// TIA Portal project "test_done_13_5" (V17)
// Vorlageprojekt für das Buch mit Zielsystem S7-1200

(* hardware
DEVICE "S71500/ET200MP station_1"  S7-1500 station
   slot 0: "Rail_0"  Rack  6ES7 590-1***0-0AA0
   slot 1: "PLC_2"  CPU 1516-3 PN/DP  6ES7 516-3AN02-0AB0  V2.8
      slot 3: "CPU display_1"  6ES7591-1BA00-0AA0
      slot 32768: "PROFINET interface_1"  X1
         slot 32769: "Port_1"  X1 P1
         slot 32770: "Port_2"  X1 P2
      slot 33024: "PROFINET interface_2"  X2
      slot 33280: "DP interface_1"  X3
      slot 34817: "Virtual CP interface port_1"  Virtual CP interface port  Virtual CP interface port
*)

// ===== PLC "PLC_2"  CPU 1516-3 PN/DP =====

VAR_GLOBAL CONSTANT   // PLC tag table "Standard-Variablentabelle"
   "Keiner" : Pip := 65535;
   "Automatische Aktualisierung" : Pip := 0;
   "TPA 1" : Pip := 1;
   "TPA 2" : Pip := 2;
   "TPA 3" : Pip := 3;
   "TPA 4" : Pip := 4;
   "TPA OB Servo" : Pip := 32768;
   "Local~MC(1)" : Hw_SubModule := 51;
   "Local~Common(1)" : Hw_SubModule := 50;
   "Local~Device(1)" : Hw_Device := 32;
   "Local~Configuration(1)" : Hw_SubModule := 33;
   "Local~Exec(1)" : Hw_SubModule := 52;
   "Local(1)" : Hw_SubModule := 49;
   "Local~PROFINET-Schnittstelle_1" : Hw_Interface := 64;
   "Local~PROFINET-Schnittstelle_1~Port_1" : Hw_Interface := 65;
   "Local~HSC_1(1)" : Hw_Hsc := 257;
   "Local~HSC_2(1)" : Hw_Hsc := 258;
   "Local~HSC_3(1)" : Hw_Hsc := 259;
   "Local~HSC_4(1)" : Hw_Hsc := 260;
   "Local~HSC_5(1)" : Hw_Hsc := 261;
   "Local~HSC_6(1)" : Hw_Hsc := 262;
   "Local~AI_2_1" : Hw_SubModule := 263;
   "Local~DI_6_DQ_4_1" : Hw_SubModule := 264;
   "Local~Pulse_1(1)" : Hw_Pwm := 265;
   "Local~Pulse_2(1)" : Hw_Pwm := 266;
   "Local~Pulse_3(1)" : Hw_Pwm := 267;
   "Local~Pulse_4(1)" : Hw_Pwm := 268;
   "OB_Main(1)" : OB_PCYCLE := 1;
END_VAR

VAR_GLOBAL   // PLC tag table "TAGS"
   "Start" AT %I0.0 : Bool;   // Nút nhấn start
   "Stop" AT %I0.1 : Bool;   // Nút nhấn stop
   "Nhap hang" AT %I0.2 : Bool;   // Nút nhấn nhập hàng
   "Xuat hang" AT %I0.3 : Bool;   // Nút nhấn xuất hàng
   "Nut tang" AT %I0.4 : Bool;   // nút nhấn tăng vị trí
   "Nut giam" AT %I0.5 : Bool;   // nút nhấn giảm vị trí
   "CB vi tri nhan hang" AT %I0.6 : Bool;   // cảm biến vị trí nhận hàng
   "CB vi tri xuat hang" AT %I0.7 : Bool;   // cảm biến vị trí xuất hàng
   "CB hang da xuat" AT %I1.0 : Bool;   // cảm biến báo hàng đã xuất
   "CB ban nang VT giua" AT %I1.1 : Bool;   // cảm biến bàn nâng ở vị trí giữa
   "CB ban nang VT phai" AT %I1.2 : Bool;   // cảm biến bàn nâng ở vị trí phải
   "CB ban nang VT Trai" AT %I1.3 : Bool;   // cảm biến bàn nâng ở vị trí trái
   "CB vi tri nhap hang" AT %I1.4 : Bool;   // cảm biến vị trí nhập hàng
   "Ban nang dang moving x" AT %I1.5 : Bool;   // bit báo bàn nâng đang di chuyển theo trục x
   "Ban nang dang moving z" AT %I1.6 : Bool;   // bit báo bàn nâng đang di chuyển theo trục z
   "Q_Den_Run" AT %Q0.0 : Bool;   // đầu ra - đèn run
   "Q_Ban_Nang_Nang_len" AT %Q0.1 : Bool;   // đầu ra - bàn nâng nâng lên
   "Q_ban nang sang phai" AT %Q0.2 : Bool;   // đầu ra - bàn nâng sang phải
   "Q ban nang sang trai" AT %Q0.3 : Bool;   // đầu ra - bàn nâng sang trái
   "Q bang tai nhap hang1" AT %Q0.4 : Bool;   // đầu ra - băng tải nhập hàng 1
   "Q bang tai nhap hang 2" AT %Q0.5 : Bool;   // đầu ra - băng tải nhập hàng 2
   "Q bang tai xuat hang 1" AT %Q0.6 : Bool;   // đầy ra - băng tải xuất hàng 1
   "Q bang tai xuat hang 2" AT %Q0.7 : Bool;   // đầu ra - băng tải xuất hàng 2
   "Cai vi tri nhap xuat hang" AT %QD34 : DInt;   // đầu ra - vị trí cần nhập xuất hàng
   "Hien thi vi tri nhap xuat hang" AT %QD38 : DInt;   // đầu ra - hiển thị vị trí đã chọn để nhập xuất hàng
END_VAR

VAR_GLOBAL   // PLC tag table "XUNG P"
   "P1" AT %M10.0 : Bool;
   "P2" AT %M10.1 : Bool;
   "P3" AT %M10.2 : Bool;
   "P4" AT %M10.3 : Bool;
   "P5" AT %M10.4 : Bool;
   "P6" AT %M10.5 : Bool;
   "P7" AT %M10.6 : Bool;
   "P8" AT %M10.7 : Bool;
   "P9" AT %M11.0 : Bool;
   "P10" AT %M11.1 : Bool;
   "P11" AT %M11.2 : Bool;
   "P12" AT %M11.3 : Bool;
   "P13" AT %M11.4 : Bool;
   "P14" AT %M11.5 : Bool;
   "P15" AT %M11.6 : Bool;
   "P16" AT %M11.7 : Bool;
   "P17" AT %M12.0 : Bool;
   "P18" AT %M12.1 : Bool;
   "P19" AT %M12.2 : Bool;
   "P20" AT %M12.3 : Bool;
END_VAR

VAR_GLOBAL   // PLC tag table "TRUNG GIAN"
   "Dang nhap hang" AT %M20.0 : Bool;
   "Dang xuat hang" AT %M20.1 : Bool;
   "Nhap hang - Buoc 1: Chay BT1,2" AT %M20.2 : Bool;
   "Nhap hang - Buoc 2: Lay hang" AT %M20.3 : Bool;
   "Nhap hang - Buoc 3: Dua hang vao vi tri" AT %M20.4 : Bool;
   "Nhap hang - Buoc 4: Ve vi tri home" AT %M20.5 : Bool;
   "TG_CB_VT_Nhan_Hang" AT %M20.6 : Bool;
   "TG_nhap_hang_buoc3" AT %M20.7 : Bool;
   "Xuat hang - Buoc 1: Di chuyen den vi tri lay" AT %M21.0 : Bool;
   "Xuat hang - Buoc 2: Lay hang" AT %M21.1 : Bool;
   "TG_xuat_hang_buoc2" AT %M21.2 : Bool;
   "Xuat hang - Buoc 3: Ve vi tri home" AT %M21.3 : Bool;
   "TG_xuat_hang_buoc3" AT %M21.4 : Bool;
   "Xuat hang - Buoc 4: BT chuyen hang di" AT %M21.5 : Bool;
   "TG_CB hang da xuat" AT %M21.6 : Bool;
   "TG_xuat_hang_buoc4" AT %M21.7 : Bool;
END_VAR

VAR_GLOBAL   // PLC tag table "TAGS MQTT"
   "MQTT_AutoEnable" AT %M30.0 : Bool;   // Luôn Enable MQTT Protocol
   "MQTT_AutoSubscribe" AT %M30.1 : Bool;
   "MQTT_Publish_Trigger" AT %M30.3 : Bool;
   "MQTT_Subscribe_Trigger" AT %M30.4 : Bool;
   "MQTT_Unsubscribe_Trigger" AT %M30.5 : Bool;
   "MQTT_Subscribe_P" AT %M30.6 : Bool;
   "Disable" AT %M30.7 : Bool;
   "Temp" AT %M31.0 : Bool;
END_VAR

// folder: Common

TYPE "typeDiagnostics"
TITLE = typeDiagnostics
// Provides a structure for detailed diagnostics
   STRUCT
      status : Word;   // Status of the block or error identification when error occurred
      subfunctionStatus : DWord;   // Status or return value of called FBs, FCs and system blocks
      stateNumber : DInt;   // State in the state machine of the block where the error occurred
   END_STRUCT;
END_TYPE

// folder: MqttClient

TYPE "MqttPublishPacket"
   STRUCT
      DUP_flag : Bool;
      QoS_level : Int;
      Retain : Bool;
      PublishTopic : String;
      PublishMessage : String;
   END_STRUCT;
END_TYPE

TYPE "MqttSubscribePacket"
   STRUCT
      TopicFilter : Array[0..9] of String;
      RequestedQoS : Array[0..9] of Byte;
   END_STRUCT;
END_TYPE

TYPE "MqttUnsubscribePacket"
   STRUCT
      TopicFilter : Array[0..9] of String;
   END_STRUCT;
END_TYPE

TYPE "MqttConnectPacket"
   STRUCT
      cleanSession : Bool := True;
      willFlag : Bool;
      willQoS_level : Int;
      willRetain : Bool;   // must be false, if Will flag is false
      passwordFlag : Bool := false;   // if true, a password is required
      userNameFlag : Bool := false;   // if true, a username is required
      keepAliveTime : Word := 10;
      clientIdentifier : String[23] := 'mqttdemo';
      willTopic : String[100] := 'myWill';
      willMessage : String[100] := 'This is my Will message';
      userName : String[20] := '';
      password : String[20] := '';
   END_STRUCT;
END_TYPE

// folder: (top level)

DATA_BLOCK "DB_WMS_Interface"   // DB17
{ S7_Optimized_Access := 'FALSE' }
VERSION : 0.1
   VAR
      Control_From_HMI : Struct
         Nhap_hang : Bool;
         Xuat_hang : Bool;
         Nut_tang : Bool;
         Nut_giam : Bool;
         Start : Bool;
         Stop : Bool;
         Cmd_Store_A01 : Bool;
         Cmd_Store_A02 : Bool;
         Cmd_Store_A03 : Bool;
         Cmd_Retrieve : Bool;
         Cmd_Reset : Bool;
      END_STRUCT;
      System_Feedback : Struct
         CB_vi_tri_nhan : Bool;
         CB_vi_tri_xuat : Bool;
         Moving_X : Bool;
         Moving_Z : Bool;
         Q_Den_Run : Bool;
      END_STRUCT;
      Warehouse_Data : Struct
         Cai_vi_tri_nhap_xuat : DInt;
         Hien_thi_vi_tri_nhap_xuat : DInt;
      END_STRUCT;
   END_VAR
BEGIN
END_DATA_BLOCK

DATA_BLOCK "MQTT_Client_DB"   // DB18
{ S7_Optimized_Access := 'TRUE' }
AUTHOR : YU_WEN_TANG
FAMILY : SLT_APC_FA
NAME : SLTAPCFA_1
VERSION : 1.0
// stored: InstanceOfName MQTT_Client
"MQTT_Client"
BEGIN
END_DATA_BLOCK

DATA_BLOCK "MqttControlPacket"   // DB19
{ S7_Optimized_Access := 'TRUE' }
VERSION : 0.1
   VAR
      ConnectPacket : "MqttConnectPacket";
      PublishPacket : "MqttPublishPacket";
      SubscribePacket : "MqttSubscribePacket";
      UnsubscribePacket : "MqttUnsubscribePacket";
   END_VAR
BEGIN
   SubscribePacket.TopicFilter[0] := 'factoryio/warehouse/cmd/system';
   PublishPacket.PublishTopic := 'factoryio/warehouse/bin_status';
   SubscribePacket.TopicFilter[1] := 'factoryio/warehouse/cmd/store';
   SubscribePacket.TopicFilter[2] := 'factoryio/warehouse/cmd/retrieve';
END_DATA_BLOCK

DATA_BLOCK "FB_Parse_MQTT_DB"   // DB20
{ S7_Optimized_Access := 'TRUE' }
VERSION : 0.1
// stored: InstanceOfName FB_Parse_MQTT
"FB_Parse_MQTT"
BEGIN
END_DATA_BLOCK

DATA_BLOCK "DB_MQTT_Control"   // DB21
{ S7_Optimized_Access := 'TRUE' }
VERSION : 0.1
   VAR
      AutoEnable : Bool := TRUE;
      PublishTrigger : Bool;
      SubscribeTrigger : Bool := false;
      SubscribeDone : Bool;
      SubscribedOK : Bool;
      MqttConnected : Bool;
      PublishCmd : Bool;
      PublishCmd_Old : Bool;
      MQTT_Subscribe_Done : Bool;
      Old_Bin_Status : Int;
      Current_Bin_Status : Int;
      PublishBusy : Bool;
      PublishDoneOld : Bool;
      PublishDoneRise : Bool;
      Current_Bin_No : Int;
      Old_Bin_No : Int;
      Current_Command : Int;
      Old_Command : Int;
   END_VAR
BEGIN
END_DATA_BLOCK

DATA_BLOCK "DB_Warehouse_Status"   // DB22
{ S7_Optimized_Access := 'TRUE' }
VERSION : 0.1
   VAR
      Bin_Empty : Bool := true;
      Bin_Occupied : Bool;
      Bin_A010101_LastEmpty : Bool;
      Bin_A010101_PublishTrigger : Bool;
      SelectedBinIndex : Int;
      SelectedBinState : Int;
   END_VAR
BEGIN
END_DATA_BLOCK

DATA_BLOCK "DB_MQTT_Warehouse"   // DB23
{ S7_Optimized_Access := 'TRUE' }
VERSION : 0.1
   VAR
      PublishTopic : String[100] := 'factoryio/warehouse/bin_status';   // topic gửi lên Node-RED
      PublishMessage : String[80];   // message ngắn
      BinIndex : Int;
      PublishRequest : Bool;   // yêu cầu publish
   END_VAR
BEGIN
END_DATA_BLOCK

// folder: System blocks/Program resources

DATA_BLOCK "IEC_Timer_0_DB"   // DB1
{ S7_Optimized_Access := 'TRUE' }
AUTHOR : Simatic
FAMILY : IEC
NAME : IEC_TMR
VERSION : 1.0
// stored: InstanceOfName IEC_TIMER
"IEC_TIMER"
BEGIN
END_DATA_BLOCK

DATA_BLOCK "IEC_Timer_0_DB_1"   // DB2
{ S7_Optimized_Access := 'TRUE' }
AUTHOR : Simatic
FAMILY : IEC
NAME : IEC_TMR
VERSION : 1.0
// stored: InstanceOfName IEC_TIMER
"IEC_TIMER"
BEGIN
END_DATA_BLOCK

DATA_BLOCK "IEC_Timer_0_DB_2"   // DB3
{ S7_Optimized_Access := 'TRUE' }
AUTHOR : Simatic
FAMILY : IEC
NAME : IEC_TMR
VERSION : 1.0
// stored: InstanceOfName IEC_TIMER
"IEC_TIMER"
BEGIN
END_DATA_BLOCK

DATA_BLOCK "IEC_Timer_0_DB_3"   // DB4
{ S7_Optimized_Access := 'TRUE' }
AUTHOR : Simatic
FAMILY : IEC
NAME : IEC_TMR
VERSION : 1.0
// stored: InstanceOfName IEC_TIMER
"IEC_TIMER"
BEGIN
END_DATA_BLOCK

DATA_BLOCK "IEC_Timer_0_DB_4"   // DB5
{ S7_Optimized_Access := 'TRUE' }
AUTHOR : Simatic
FAMILY : IEC
NAME : IEC_TMR
VERSION : 1.0
// stored: InstanceOfName IEC_TIMER
"IEC_TIMER"
BEGIN
END_DATA_BLOCK

DATA_BLOCK "IEC_Timer_0_DB_5"   // DB6
{ S7_Optimized_Access := 'TRUE' }
AUTHOR : Simatic
FAMILY : IEC
NAME : IEC_TMR
VERSION : 1.0
// stored: InstanceOfName IEC_TIMER
"IEC_TIMER"
BEGIN
END_DATA_BLOCK

DATA_BLOCK "IEC_Timer_0_DB_6"   // DB7
{ S7_Optimized_Access := 'TRUE' }
AUTHOR : Simatic
FAMILY : IEC
NAME : IEC_TMR
VERSION : 1.0
// stored: InstanceOfName IEC_TIMER
"IEC_TIMER"
BEGIN
END_DATA_BLOCK

DATA_BLOCK "IEC_Timer_0_DB_7"   // DB8
{ S7_Optimized_Access := 'TRUE' }
AUTHOR : Simatic
FAMILY : IEC
NAME : IEC_TMR
VERSION : 1.0
// stored: InstanceOfName IEC_TIMER
"IEC_TIMER"
BEGIN
END_DATA_BLOCK

DATA_BLOCK "IEC_Timer_0_DB_8"   // DB9
{ S7_Optimized_Access := 'TRUE' }
AUTHOR : Simatic
FAMILY : IEC
NAME : IEC_TMR
VERSION : 1.0
// stored: InstanceOfName IEC_TIMER
"IEC_TIMER"
BEGIN
END_DATA_BLOCK

DATA_BLOCK "IEC_Timer_0_DB_9"   // DB10
{ S7_Optimized_Access := 'TRUE' }
AUTHOR : Simatic
FAMILY : IEC
NAME : IEC_TMR
VERSION : 1.0
// stored: InstanceOfName IEC_TIMER
"IEC_TIMER"
BEGIN
END_DATA_BLOCK

DATA_BLOCK "IEC_Timer_0_DB_10"   // DB11
{ S7_Optimized_Access := 'TRUE' }
AUTHOR : Simatic
FAMILY : IEC
NAME : IEC_TMR
VERSION : 1.0
// stored: InstanceOfName IEC_TIMER
"IEC_TIMER"
BEGIN
END_DATA_BLOCK

DATA_BLOCK "IEC_Timer_0_DB_11"   // DB12
{ S7_Optimized_Access := 'TRUE' }
AUTHOR : Simatic
FAMILY : IEC
NAME : IEC_TMR
VERSION : 1.0
// stored: InstanceOfName IEC_TIMER
"IEC_TIMER"
BEGIN
END_DATA_BLOCK

DATA_BLOCK "IEC_Timer_0_DB_12"   // DB13
{ S7_Optimized_Access := 'TRUE' }
AUTHOR : Simatic
FAMILY : IEC
NAME : IEC_TMR
VERSION : 1.0
// stored: InstanceOfName IEC_TIMER
"IEC_TIMER"
BEGIN
END_DATA_BLOCK

DATA_BLOCK "IEC_Timer_0_DB_13"   // DB14
{ S7_Optimized_Access := 'TRUE' }
AUTHOR : Simatic
FAMILY : IEC
NAME : IEC_TMR
VERSION : 1.0
// stored: InstanceOfName IEC_TIMER
"IEC_TIMER"
BEGIN
END_DATA_BLOCK

DATA_BLOCK "IEC_Timer_0_DB_14"   // DB15
{ S7_Optimized_Access := 'TRUE' }
AUTHOR : Simatic
FAMILY : IEC
NAME : IEC_TMR
VERSION : 1.0
// stored: InstanceOfName IEC_TIMER
"IEC_TIMER"
BEGIN
END_DATA_BLOCK

DATA_BLOCK "IEC_Timer_0_DB_15"   // DB16
{ S7_Optimized_Access := 'TRUE' }
AUTHOR : Simatic
FAMILY : IEC
NAME : IEC_TMR
VERSION : 1.0
// stored: InstanceOfName IEC_TIMER
"IEC_TIMER"
BEGIN
END_DATA_BLOCK

// folder: (top level)

FUNCTION_BLOCK "FB_Parse_MQTT"   // FB1, SCL
{ S7_Optimized_Access := 'TRUE' }
VERSION : 0.1
   VAR_INPUT
      ReceivedMessage : String;
      ReceivedTopic : String;
   END_VAR
   VAR_OUTPUT
      Nhap_hang : Bool;
      Xuat_hang : Bool;
      Vi_tri : DInt;
      Start : Bool;
      Stop : Bool;
   END_VAR
   VAR
      LastMessage : String;
      LastTopic : String;
   END_VAR
BEGIN
   #Start := FALSE;
   #Stop := FALSE;
   #Nhap_hang := FALSE;
   #Xuat_hang := FALSE;

   IF (#ReceivedTopic <> #LastTopic) OR (#ReceivedMessage <> #LastMessage) THEN

       IF #ReceivedTopic = 'factoryio/warehouse/cmd/system' THEN
           IF #ReceivedMessage = 'START' THEN
               #Start := TRUE;
           END_IF;

           IF #ReceivedMessage = 'STOP' THEN
               #Stop := TRUE;
           END_IF;
       END_IF;

       IF #ReceivedTopic = 'factoryio/warehouse/cmd/store' THEN
           #Nhap_hang := TRUE;
           #Vi_tri := STRING_TO_DINT(#ReceivedMessage);
       END_IF;

       IF #ReceivedTopic = 'factoryio/warehouse/cmd/retrieve' THEN
           #Xuat_hang := TRUE;
           #Vi_tri := STRING_TO_DINT(#ReceivedMessage);
       END_IF;

       #LastTopic := #ReceivedTopic;
       #LastMessage := #ReceivedMessage;

   END_IF;
END_FUNCTION_BLOCK

FUNCTION "FC_Build_Bin_MQTT_Message" : Void   // FC1, SCL
{ S7_Optimized_Access := 'TRUE' }
VERSION : 0.1
   VAR_INPUT
      BinIndex : Int;
      State : Int;
   END_VAR
   VAR_OUTPUT
      MQTT_Message : String;
   END_VAR
BEGIN
   #MQTT_Message := CONCAT(IN1 := INT_TO_STRING(#BinIndex), IN2 := ',');
   #MQTT_Message := CONCAT(IN1 := #MQTT_Message, IN2 := INT_TO_STRING(#State));
END_FUNCTION

FUNCTION "MHJ-PLC-Lab-Function-S71200" : Void   // FC9000, SCL
{ S7_Optimized_Access := 'TRUE' }
VERSION : 0.1
   VAR_TEMP
      rdTimeReturn : Int;
      outputTime : DTL;
      SyncVal : Byte;
      forVal : Int;
      forVal_2 : Int;
      Value : Byte;
   END_VAR
   VAR CONSTANT
      CompVal : Byte := 16#34;
      Value_01 : Byte := 16#11;
      Value_01_DW : DWord := 16#A165_D992;
      Value_02_DW : DWord := 16#58BE_4401;
   END_VAR
BEGIN

   #Value:=PEEK(area := 16#82,
        dbNumber := 0,
        byteOffset := 511);
   #Value := #Value + 1;

   POKE(area := 16#82,
        dbNumber := 0,
        byteOffset := 511,
        value := #Value);

   POKE(area:=16#81,
        dbNumber:=0,
        byteOffset:=1016,
        value:=#Value_01_DW);
   POKE(area := 16#81,
        dbNumber := 0,
        byteOffset := 1020,
        value := #Value_02_DW);

   POKE(area := 16#81,
        dbNumber := 0,
        byteOffset := 511,
        value := B#16#00);

   FOR #forVal := 0 TO 120 DO
       FOR #forVal_2:=0 TO 10 DO
           #rdTimeReturn:=RD_SYS_T(#outputTime);
           #rdTimeReturn := WR_SYS_T(#outputTime);
           #rdTimeReturn := RD_SYS_T(#outputTime);
           #rdTimeReturn := WR_SYS_T(#outputTime);
       END_FOR;
       #SyncVal:= PEEK(area := 16#81,
                      dbNumber := 0,
                      byteOffset := 511);
       IF #SyncVal = #CompVal THEN
          GOTO M_1;
       END_IF;
   END_FOR;
   RETURN;

   M_1:
   POKE(area := 16#81,
        dbNumber := 0,
        byteOffset := 511,
        value := B#16#0);
END_FUNCTION

ORGANIZATION_BLOCK "Main"   // OB1, LAD, ProgramCycle
TITLE = "Main Program Sweep (Cycle)"
{ S7_Optimized_Access := 'TRUE' }
VERSION : 0.1
   VAR_INPUT
      Initial_Call : Bool;   // Initial call of this OB
      Remanence : Bool;   // =True, if remanent data are available
   END_VAR
   VAR_TEMP   // added for the SCL form of the ladder/FBD networks
      _w1 : Bool;
      _w2 : Bool;
      _w3 : Bool;
      _w4 : Bool;
   END_VAR
BEGIN

REGION Network 1: Konnektierungsbaustein für PLC-Lab
   // Im Netzwerk 1 wird der Konnektierungsbaustein für PLC-Lab aufgerufen.
   // Dieser Aufruf darf nicht entfernt werden!
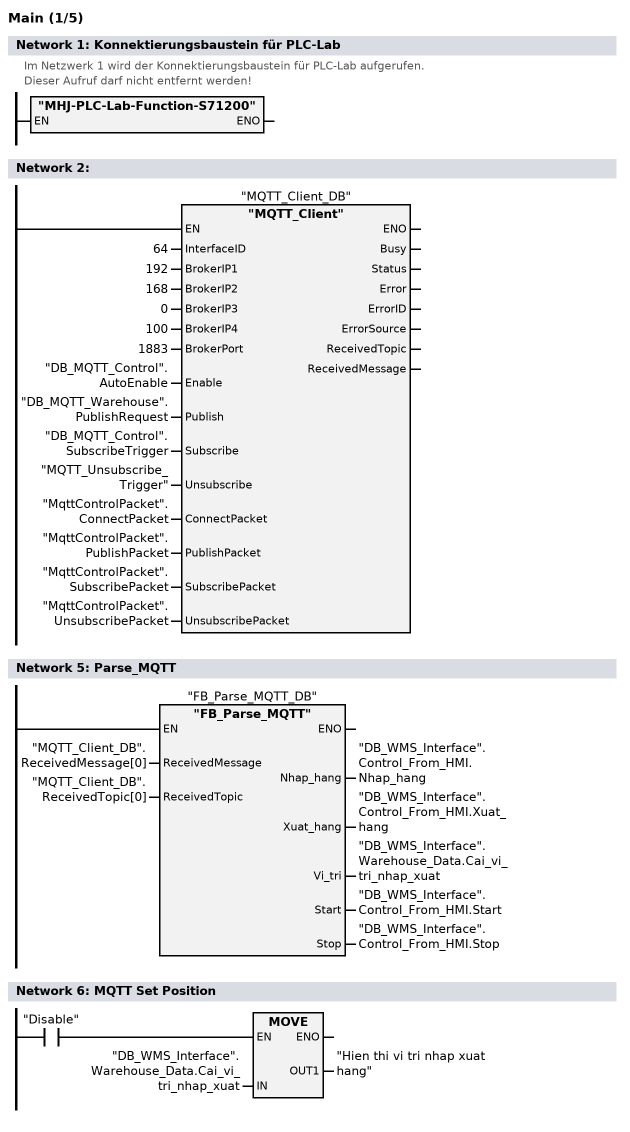
   RUNG wire#powerrail
      "MHJ-PLC-Lab-Function-S71200"()
   END_RUNG
   // the same network as SCL:
   "MHJ-PLC-Lab-Function-S71200"();
END_REGION

REGION Network 2
   RUNG wire#powerrail
      "MQTT_Client_DB"(InterfaceID := 64, BrokerIP1 := 192, BrokerIP2 := 168, BrokerIP3 := 0, BrokerIP4 := 100, BrokerPort := 1883, Enable := "DB_MQTT_Control".AutoEnable, Publish := "DB_MQTT_Warehouse".PublishRequest, Subscribe := "DB_MQTT_Control".SubscribeTrigger, Unsubscribe := "MQTT_Unsubscribe_Trigger", ConnectPacket := "MqttControlPacket".ConnectPacket, PublishPacket := "MqttControlPacket".PublishPacket, SubscribePacket := "MqttControlPacket".SubscribePacket, UnsubscribePacket := "MqttControlPacket".UnsubscribePacket, Busy =>, Status =>, Error =>, ErrorID =>, ErrorSource =>, ReceivedTopic =>, ReceivedMessage =>)
   END_RUNG
   // the same network as SCL:
   "MQTT_Client_DB"(InterfaceID := 64,   // "MQTT_Client"
                    BrokerIP1 := 192,
                    BrokerIP2 := 168,
                    BrokerIP3 := 0,
                    BrokerIP4 := 100,
                    BrokerPort := 1883,
                    Enable := "DB_MQTT_Control".AutoEnable,
                    Publish := "DB_MQTT_Warehouse".PublishRequest,
                    Subscribe := "DB_MQTT_Control".SubscribeTrigger,
                    Unsubscribe := "MQTT_Unsubscribe_Trigger",
                    ConnectPacket := "MqttControlPacket".ConnectPacket,
                    PublishPacket := "MqttControlPacket".PublishPacket,
                    SubscribePacket := "MqttControlPacket".SubscribePacket,
                    UnsubscribePacket := "MqttControlPacket".UnsubscribePacket);
END_REGION

REGION Network 3 (SCL)
   IF "MQTT_Client_DB".Status.%X1 AND NOT "DB_MQTT_Control".SubscribeDone THEN
       "DB_MQTT_Control".SubscribeTrigger := TRUE;
   END_IF;

   IF "MQTT_Client_DB".Status.%X3 THEN
       "DB_MQTT_Control".SubscribeTrigger := FALSE;
       "DB_MQTT_Control".SubscribeDone := TRUE;
   END_IF;
END_REGION

REGION Network 4 (SCL)
   // Lấy số bin hiện tại
   "DB_MQTT_Control".Current_Bin_No :=
   "DB_WMS_Interface".Warehouse_Data.Cai_vi_tri_nhap_xuat;


   // Xác định lệnh hiện tại
   // 1 = STORE, 2 = RETRIEVE, 0 = không có lệnh
   IF "Dang nhap hang" THEN

       "DB_MQTT_Control".Current_Command := 1;

   ELSIF "Dang xuat hang" THEN

       "DB_MQTT_Control".Current_Command := 2;

   ELSE

       "DB_MQTT_Control".Current_Command := 0;

   END_IF;


   // Bắt cạnh lên của Publish Done
   "DB_MQTT_Control".PublishDoneRise :=
   "MQTT_Client_DB".Status.%X2
   AND NOT "DB_MQTT_Control".PublishDoneOld;

   "DB_MQTT_Control".PublishDoneOld :=
   "MQTT_Client_DB".Status.%X2;


   // Khi MQTT đã connected,
   // chưa publish bận,
   // command khác 0,
   // và bin hoặc command thay đổi
   // thì tự publish
   IF "MQTT_Client_DB".Status.%X1
       AND NOT "DB_MQTT_Control".PublishBusy
       AND "DB_MQTT_Control".Current_Command <> 0
       AND (
       "DB_MQTT_Control".Current_Bin_No <> "DB_MQTT_Control".Old_Bin_No
       OR
       "DB_MQTT_Control".Current_Command <> "DB_MQTT_Control".Old_Command
       )
   THEN

       "DB_MQTT_Warehouse".PublishRequest := TRUE;

       "DB_MQTT_Control".PublishBusy := TRUE;

       "DB_MQTT_Control".Old_Bin_No :=
       "DB_MQTT_Control".Current_Bin_No;

       "DB_MQTT_Control".Old_Command :=
       "DB_MQTT_Control".Current_Command;

   END_IF;


   // Khi publish xong thì tắt PublishRequest
   IF "DB_MQTT_Control".PublishBusy
       AND "DB_MQTT_Control".PublishDoneRise
   THEN

       "DB_MQTT_Warehouse".PublishRequest := FALSE;

       "DB_MQTT_Control".PublishBusy := FALSE;

   END_IF;
END_REGION

REGION Network 5: Parse_MQTT
   RUNG wire#powerrail
      "FB_Parse_MQTT_DB"(ReceivedMessage := "MQTT_Client_DB".ReceivedMessage[0], ReceivedTopic := "MQTT_Client_DB".ReceivedTopic[0], Nhap_hang => "DB_WMS_Interface".Control_From_HMI.Nhap_hang, Xuat_hang => "DB_WMS_Interface".Control_From_HMI.Xuat_hang, Vi_tri => "DB_WMS_Interface".Warehouse_Data.Cai_vi_tri_nhap_xuat, Start => "DB_WMS_Interface".Control_From_HMI.Start, Stop => "DB_WMS_Interface".Control_From_HMI.Stop)
   END_RUNG
   // the same network as SCL:
   "FB_Parse_MQTT_DB"(ReceivedMessage := "MQTT_Client_DB".ReceivedMessage[0],   // "FB_Parse_MQTT"
                      ReceivedTopic := "MQTT_Client_DB".ReceivedTopic[0],
                      Nhap_hang => "DB_WMS_Interface".Control_From_HMI.Nhap_hang,
                      Xuat_hang => "DB_WMS_Interface".Control_From_HMI.Xuat_hang,
                      Vi_tri => "DB_WMS_Interface".Warehouse_Data.Cai_vi_tri_nhap_xuat,
                      Start => "DB_WMS_Interface".Control_From_HMI.Start,
                      Stop => "DB_WMS_Interface".Control_From_HMI.Stop);
END_REGION

REGION Network 6: MQTT Set Position
   RUNG wire#powerrail
      Contact( "Disable" )
      Move(in := "DB_WMS_Interface".Warehouse_Data.Cai_vi_tri_nhap_xuat, out1 => "Hien thi vi tri nhap xuat hang")
   END_RUNG
   // the same network as SCL:
   IF "Disable" THEN
       "Hien thi vi tri nhap xuat hang" := "DB_WMS_Interface".Warehouse_Data.Cai_vi_tri_nhap_xuat;
   END_IF;
END_REGION

REGION Network 7: Ihr Programm / Điều khiển hệ thống
   // Schreiben Sie ab Netzwerk 2 Ihr Programm
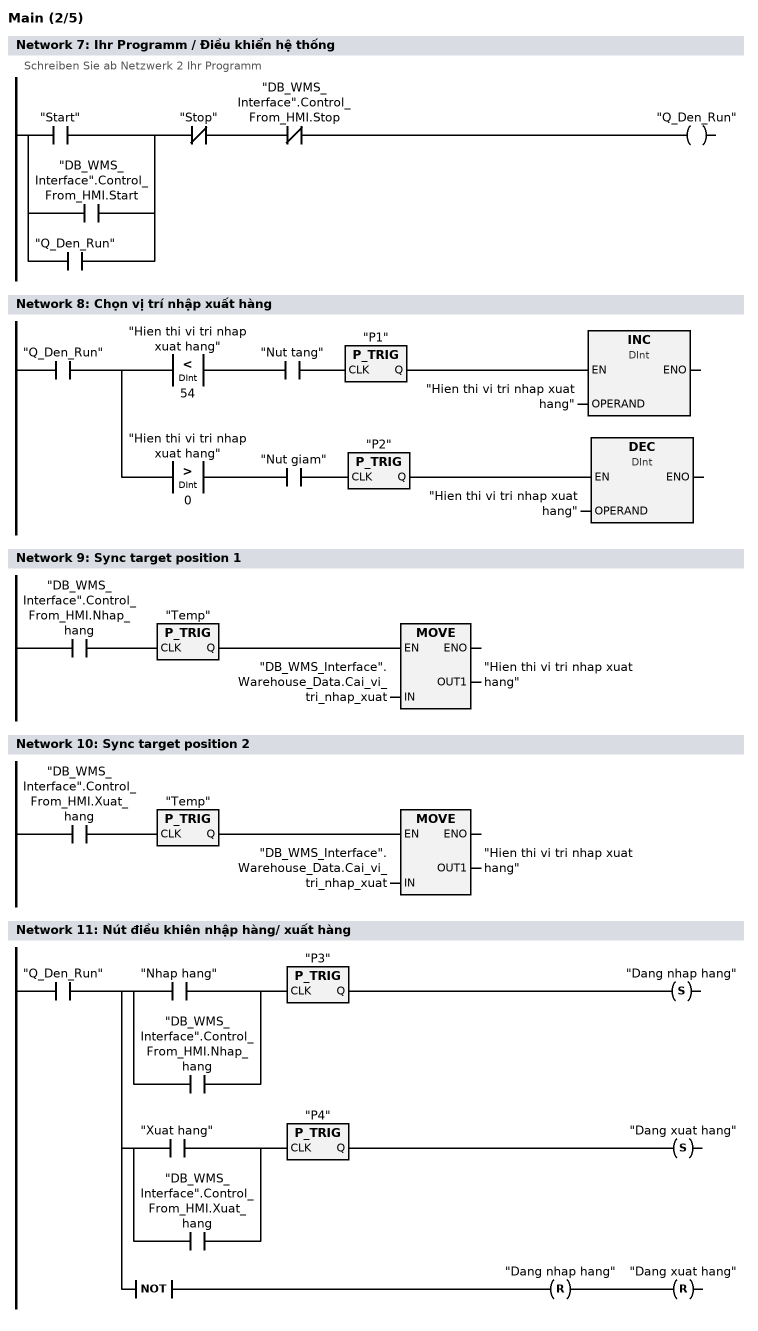
   RUNG wire#powerrail
      Contact( "Start" )
      wire#w1
      I_Contact( "Stop" )
      I_Contact( "DB_WMS_Interface".Control_From_HMI.Stop )
      Coil( "Q_Den_Run" )
   END_RUNG
   RUNG wire#powerrail
      Contact( "DB_WMS_Interface".Control_From_HMI.Start )
   END_RUNG wire#w1
   RUNG wire#powerrail
      Contact( "Q_Den_Run" )
   END_RUNG wire#w1
   // the same network as SCL:
   "Q_Den_Run" := ("Start" OR "DB_WMS_Interface".Control_From_HMI.Start OR "Q_Den_Run") AND NOT "Stop" AND NOT "DB_WMS_Interface".Control_From_HMI.Stop;
END_REGION

REGION Network 8: Chọn vị trí nhập xuất hàng
   RUNG wire#powerrail
      Contact( "Q_Den_Run" )
      wire#w1
      { S7_Templates := "SrcType := DInt" } LT_Contact(in1 := "Hien thi vi tri nhap xuat hang", in2 := 54)
      Contact( "Nut tang" )
      P_Trig( "P1" )
      { S7_Templates := "DestType := DInt" } Inc( "Hien thi vi tri nhap xuat hang" )
   END_RUNG
   RUNG wire#w1
      { S7_Templates := "SrcType := DInt" } GT_Contact(in1 := "Hien thi vi tri nhap xuat hang", in2 := 0)
      Contact( "Nut giam" )
      P_Trig( "P2" )
      { S7_Templates := "DestType := DInt" } Dec( "Hien thi vi tri nhap xuat hang" )
   END_RUNG
   // the same network as SCL:
   #_w1 := "Q_Den_Run" AND ("Hien thi vi tri nhap xuat hang" < 54) AND "Nut tang";
   #_w2 := #_w1 AND NOT "P1";   // rising edge
   "P1" := #_w1;
   IF #_w2 THEN "Hien thi vi tri nhap xuat hang" := "Hien thi vi tri nhap xuat hang" + 1; END_IF;
   #_w3 := "Q_Den_Run" AND ("Hien thi vi tri nhap xuat hang" > 0) AND "Nut giam";
   #_w4 := #_w3 AND NOT "P2";   // rising edge
   "P2" := #_w3;
   IF #_w4 THEN "Hien thi vi tri nhap xuat hang" := "Hien thi vi tri nhap xuat hang" - 1; END_IF;
END_REGION

REGION Network 9: Sync target position 1
   RUNG wire#powerrail
      Contact( "DB_WMS_Interface".Control_From_HMI.Nhap_hang )
      P_Trig( "Temp" )
      Move(in := "DB_WMS_Interface".Warehouse_Data.Cai_vi_tri_nhap_xuat, out1 => "Hien thi vi tri nhap xuat hang")
   END_RUNG
   // the same network as SCL:
   #_w1 := "DB_WMS_Interface".Control_From_HMI.Nhap_hang AND NOT "Temp";   // rising edge
   "Temp" := "DB_WMS_Interface".Control_From_HMI.Nhap_hang;
   IF #_w1 THEN
       "Hien thi vi tri nhap xuat hang" := "DB_WMS_Interface".Warehouse_Data.Cai_vi_tri_nhap_xuat;
   END_IF;
END_REGION

REGION Network 10: Sync target position 2
   RUNG wire#powerrail
      Contact( "DB_WMS_Interface".Control_From_HMI.Xuat_hang )
      P_Trig( "Temp" )
      Move(in := "DB_WMS_Interface".Warehouse_Data.Cai_vi_tri_nhap_xuat, out1 => "Hien thi vi tri nhap xuat hang")
   END_RUNG
   // the same network as SCL:
   #_w1 := "DB_WMS_Interface".Control_From_HMI.Xuat_hang AND NOT "Temp";   // rising edge
   "Temp" := "DB_WMS_Interface".Control_From_HMI.Xuat_hang;
   IF #_w1 THEN
       "Hien thi vi tri nhap xuat hang" := "DB_WMS_Interface".Warehouse_Data.Cai_vi_tri_nhap_xuat;
   END_IF;
END_REGION

REGION Network 11: Nút điều khiên nhập hàng/ xuất hàng
   RUNG wire#powerrail
      Contact( "Q_Den_Run" )
      wire#w1
      Contact( "Nhap hang" )
      wire#w2
      P_Trig( "P3" )
      S_Coil( "Dang nhap hang" )
   END_RUNG
   RUNG wire#w1
      Contact( "DB_WMS_Interface".Control_From_HMI.Nhap_hang )
   END_RUNG wire#w2
   RUNG wire#w1
      Contact( "Xuat hang" )
      wire#w3
      P_Trig( "P4" )
      S_Coil( "Dang xuat hang" )
   END_RUNG
   RUNG wire#w1
      Contact( "DB_WMS_Interface".Control_From_HMI.Xuat_hang )
   END_RUNG wire#w3
   RUNG wire#w1
      Not()
      R_Coil( "Dang nhap hang" )
      R_Coil( "Dang xuat hang" )
   END_RUNG
   // the same network as SCL:
   #_w1 := "Q_Den_Run" AND ("Nhap hang" OR "DB_WMS_Interface".Control_From_HMI.Nhap_hang);
   #_w2 := #_w1 AND NOT "P3";   // rising edge
   "P3" := #_w1;
   IF #_w2 THEN "Dang nhap hang" := TRUE; END_IF;
   #_w3 := "Q_Den_Run" AND ("Xuat hang" OR "DB_WMS_Interface".Control_From_HMI.Xuat_hang);
   #_w4 := #_w3 AND NOT "P4";   // rising edge
   "P4" := #_w3;
   IF #_w4 THEN "Dang xuat hang" := TRUE; END_IF;
   IF NOT "Q_Den_Run" THEN
       "Dang nhap hang" := FALSE;
       "Dang xuat hang" := FALSE;
   END_IF;
END_REGION

REGION Network 12: Đang nhập hàng - bước 1
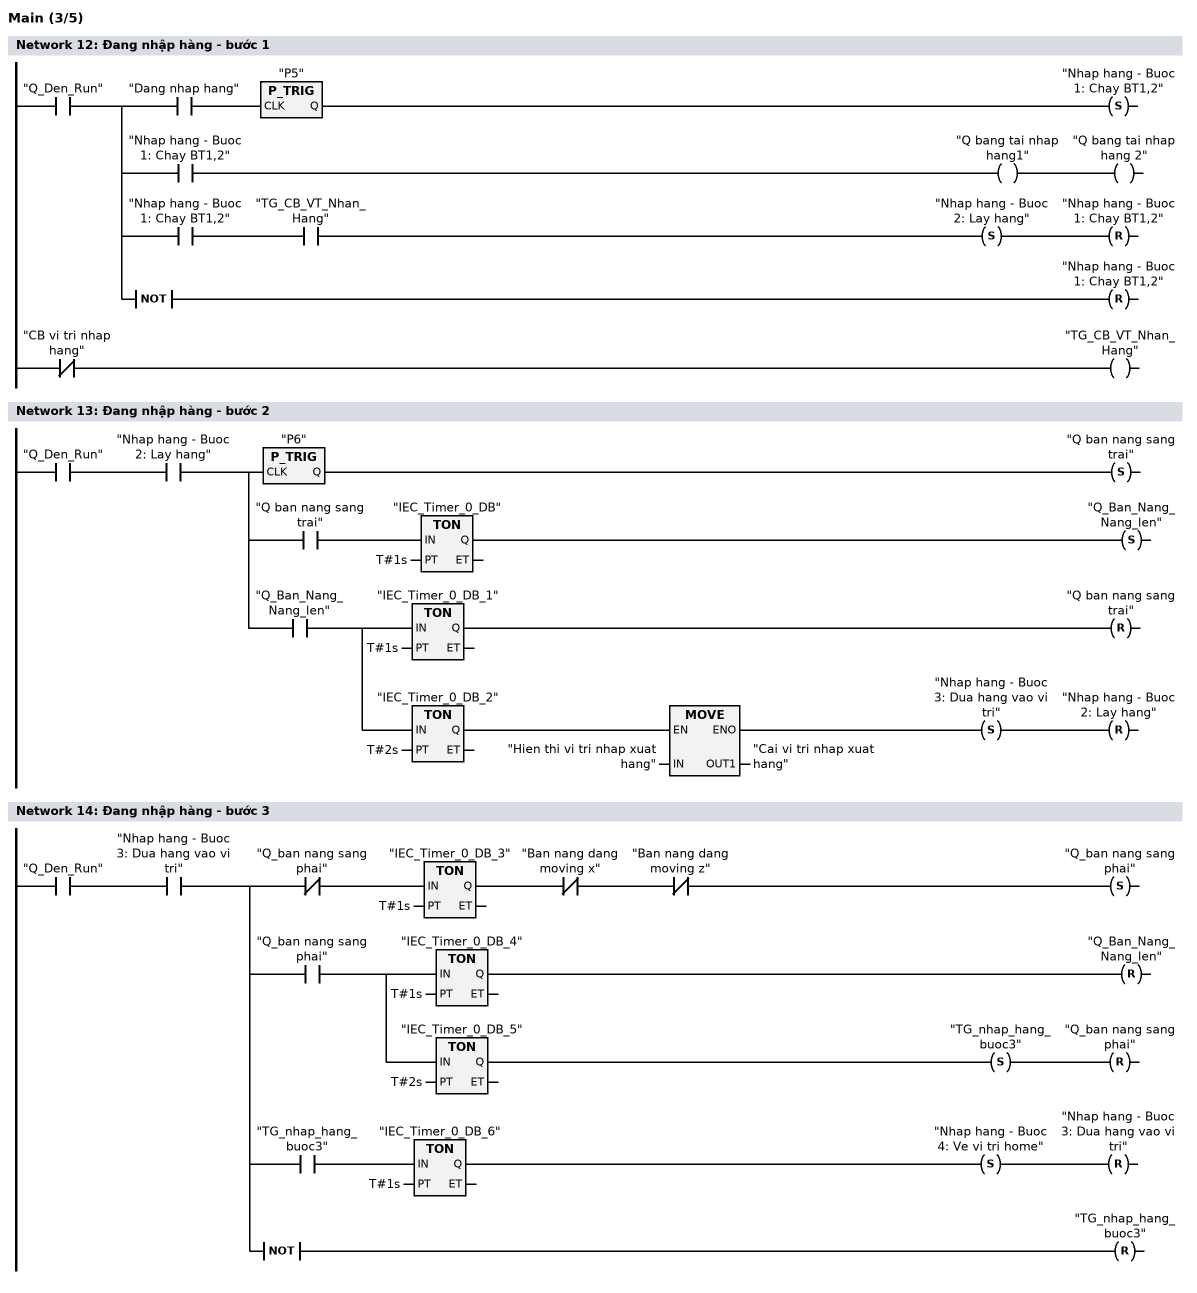
   RUNG wire#powerrail
      Contact( "Q_Den_Run" )
      wire#w1
      Contact( "Dang nhap hang" )
      P_Trig( "P5" )
      S_Coil( "Nhap hang - Buoc 1: Chay BT1,2" )
   END_RUNG
   RUNG wire#w1
      Contact( "Nhap hang - Buoc 1: Chay BT1,2" )
      Coil( "Q bang tai nhap hang1" )
      Coil( "Q bang tai nhap hang 2" )
   END_RUNG
   RUNG wire#w1
      Contact( "Nhap hang - Buoc 1: Chay BT1,2" )
      Contact( "TG_CB_VT_Nhan_Hang" )
      S_Coil( "Nhap hang - Buoc 2: Lay hang" )
      R_Coil( "Nhap hang - Buoc 1: Chay BT1,2" )
   END_RUNG
   RUNG wire#w1
      Not()
      R_Coil( "Nhap hang - Buoc 1: Chay BT1,2" )
   END_RUNG
   RUNG wire#powerrail
      I_Contact( "CB vi tri nhap hang" )
      Coil( "TG_CB_VT_Nhan_Hang" )
   END_RUNG
   // the same network as SCL:
   #_w1 := "Q_Den_Run" AND "Dang nhap hang";
   #_w2 := #_w1 AND NOT "P5";   // rising edge
   "P5" := #_w1;
   IF #_w2 THEN "Nhap hang - Buoc 1: Chay BT1,2" := TRUE; END_IF;
   "Q bang tai nhap hang1" := "Q_Den_Run" AND "Nhap hang - Buoc 1: Chay BT1,2";
   "Q bang tai nhap hang 2" := "Q bang tai nhap hang1";
   IF "Q_Den_Run" AND "Nhap hang - Buoc 1: Chay BT1,2" AND "TG_CB_VT_Nhan_Hang" THEN
       "Nhap hang - Buoc 2: Lay hang" := TRUE;
       "Nhap hang - Buoc 1: Chay BT1,2" := FALSE;
   END_IF;
   IF NOT "Q_Den_Run" THEN "Nhap hang - Buoc 1: Chay BT1,2" := FALSE; END_IF;
   "TG_CB_VT_Nhan_Hang" := NOT "CB vi tri nhap hang";
END_REGION

REGION Network 13: Đang nhập hàng - bước 2
   #_w1 := "Q_Den_Run" AND "Nhap hang - Buoc 2: Lay hang";
   #_w2 := #_w1 AND NOT "P6";   // rising edge
   "P6" := #_w1;
   IF #_w2 THEN "Q ban nang sang trai" := TRUE; END_IF;
   "IEC_Timer_0_DB".TON(IN := #_w1 AND "Q ban nang sang trai", PT := T#1s);
   IF "IEC_Timer_0_DB".Q THEN "Q_Ban_Nang_Nang_len" := TRUE; END_IF;
   #_w3 := #_w1 AND "Q_Ban_Nang_Nang_len";
   "IEC_Timer_0_DB_1".TON(IN := #_w3, PT := T#1s);
   IF "IEC_Timer_0_DB_1".Q THEN "Q ban nang sang trai" := FALSE; END_IF;
   "IEC_Timer_0_DB_2".TON(IN := #_w3, PT := T#2s);
   IF "IEC_Timer_0_DB_2".Q THEN
       "Cai vi tri nhap xuat hang" := "Hien thi vi tri nhap xuat hang";
       "Nhap hang - Buoc 3: Dua hang vao vi tri" := TRUE;
       "Nhap hang - Buoc 2: Lay hang" := FALSE;
   END_IF;
END_REGION

REGION Network 14: Đang nhập hàng - bước 3
   #_w1 := "Q_Den_Run" AND "Nhap hang - Buoc 3: Dua hang vao vi tri";
   "IEC_Timer_0_DB_3".TON(IN := #_w1 AND NOT "Q_ban nang sang phai", PT := T#1s);
   IF "IEC_Timer_0_DB_3".Q AND NOT "Ban nang dang moving x" AND NOT "Ban nang dang moving z" THEN
       "Q_ban nang sang phai" := TRUE;
   END_IF;
   #_w2 := #_w1 AND "Q_ban nang sang phai";
   "IEC_Timer_0_DB_4".TON(IN := #_w2, PT := T#1s);
   IF "IEC_Timer_0_DB_4".Q THEN "Q_Ban_Nang_Nang_len" := FALSE; END_IF;
   "IEC_Timer_0_DB_5".TON(IN := #_w2, PT := T#2s);
   IF "IEC_Timer_0_DB_5".Q THEN
       "TG_nhap_hang_buoc3" := TRUE;
       "Q_ban nang sang phai" := FALSE;
   END_IF;
   "IEC_Timer_0_DB_6".TON(IN := #_w1 AND "TG_nhap_hang_buoc3", PT := T#1s);
   IF "IEC_Timer_0_DB_6".Q THEN
       "Nhap hang - Buoc 4: Ve vi tri home" := TRUE;
       "Nhap hang - Buoc 3: Dua hang vao vi tri" := FALSE;
   END_IF;
   IF NOT #_w1 THEN "TG_nhap_hang_buoc3" := FALSE; END_IF;
END_REGION

REGION Network 15: Đang nhập hàng - bước 4
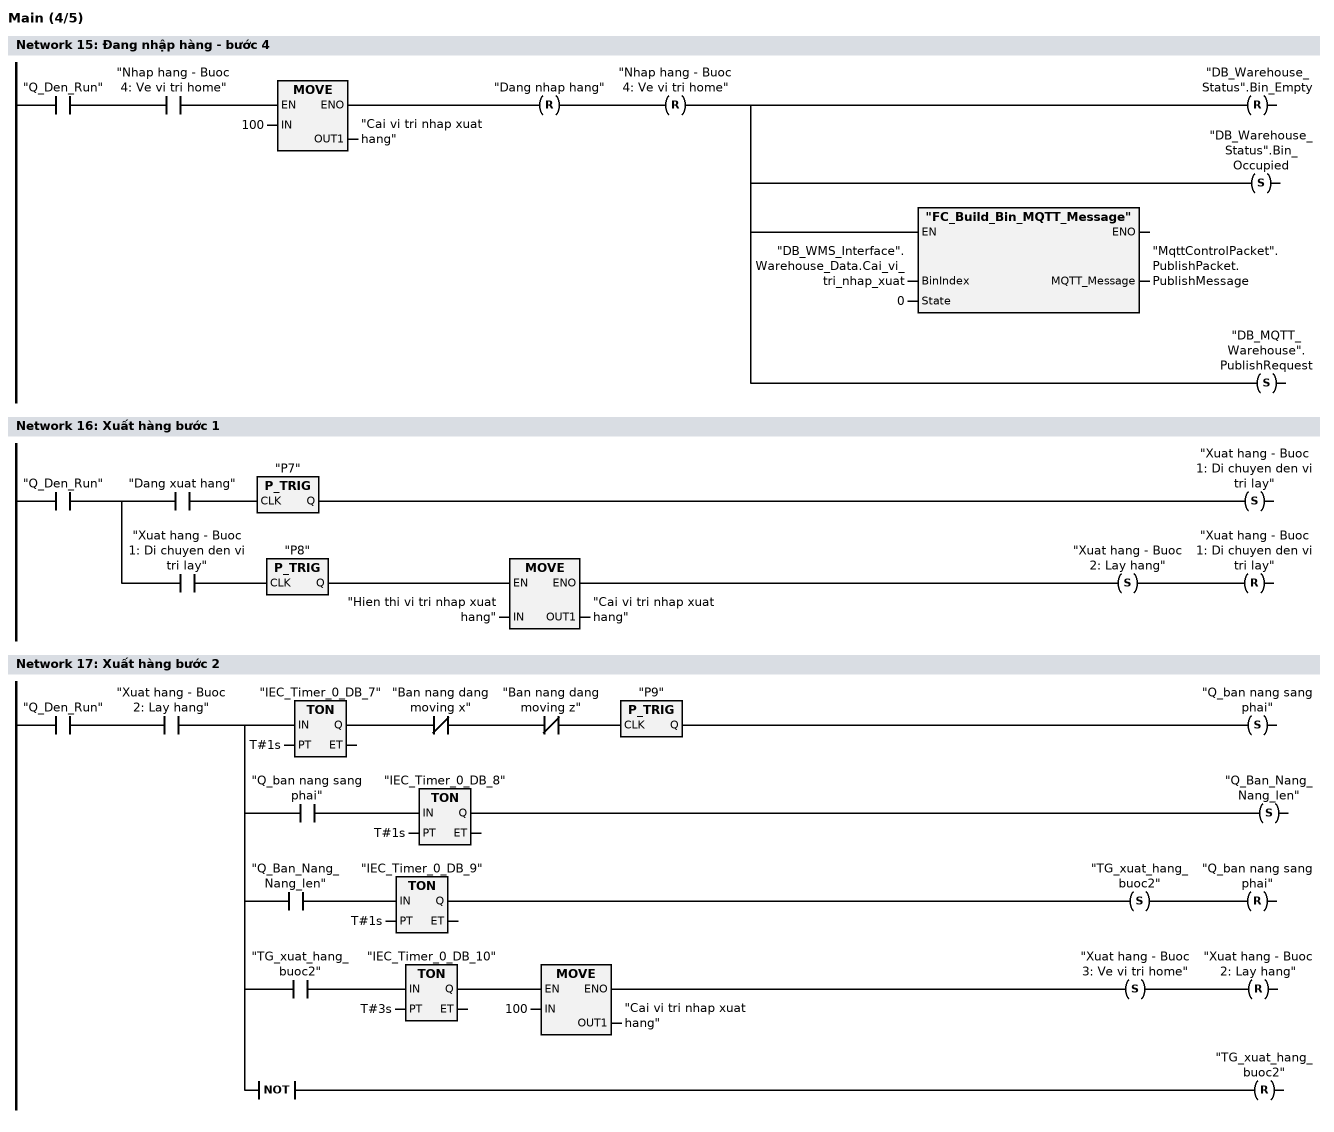
   RUNG wire#powerrail
      Contact( "Q_Den_Run" )
      Contact( "Nhap hang - Buoc 4: Ve vi tri home" )
      Move(in := 100, out1 => "Cai vi tri nhap xuat hang")
      R_Coil( "Dang nhap hang" )
      R_Coil( "Nhap hang - Buoc 4: Ve vi tri home" )
      wire#w1
      R_Coil( "DB_Warehouse_Status".Bin_Empty )
   END_RUNG
   RUNG wire#w1
      S_Coil( "DB_Warehouse_Status".Bin_Occupied )
   END_RUNG
   RUNG wire#w1
      "FC_Build_Bin_MQTT_Message"(BinIndex := "DB_WMS_Interface".Warehouse_Data.Cai_vi_tri_nhap_xuat, State := 0, MQTT_Message => "MqttControlPacket".PublishPacket.PublishMessage)
   END_RUNG
   RUNG wire#w1
      S_Coil( "DB_MQTT_Warehouse".PublishRequest )
   END_RUNG
   // the same network as SCL:
   IF "Q_Den_Run" AND "Nhap hang - Buoc 4: Ve vi tri home" THEN
       "Cai vi tri nhap xuat hang" := 100;
       "Dang nhap hang" := FALSE;
   END_IF;
   #_w1 := "Q_Den_Run" AND "Nhap hang - Buoc 4: Ve vi tri home";
   IF #_w1 THEN
       "Nhap hang - Buoc 4: Ve vi tri home" := FALSE;
       "DB_Warehouse_Status".Bin_Empty := FALSE;
       "DB_Warehouse_Status".Bin_Occupied := TRUE;
       "FC_Build_Bin_MQTT_Message"(BinIndex := "DB_WMS_Interface".Warehouse_Data.Cai_vi_tri_nhap_xuat,
                               State := 0,
                               MQTT_Message => "MqttControlPacket".PublishPacket.PublishMessage);
       "DB_MQTT_Warehouse".PublishRequest := TRUE;
   END_IF;
END_REGION

REGION Network 16: Xuất hàng bước 1
   RUNG wire#powerrail
      Contact( "Q_Den_Run" )
      wire#w1
      Contact( "Dang xuat hang" )
      P_Trig( "P7" )
      S_Coil( "Xuat hang - Buoc 1: Di chuyen den vi tri lay" )
   END_RUNG
   RUNG wire#w1
      Contact( "Xuat hang - Buoc 1: Di chuyen den vi tri lay" )
      P_Trig( "P8" )
      Move(in := "Hien thi vi tri nhap xuat hang", out1 => "Cai vi tri nhap xuat hang")
      S_Coil( "Xuat hang - Buoc 2: Lay hang" )
      R_Coil( "Xuat hang - Buoc 1: Di chuyen den vi tri lay" )
   END_RUNG
   // the same network as SCL:
   #_w1 := "Q_Den_Run" AND "Dang xuat hang";
   #_w2 := #_w1 AND NOT "P7";   // rising edge
   "P7" := #_w1;
   IF #_w2 THEN "Xuat hang - Buoc 1: Di chuyen den vi tri lay" := TRUE; END_IF;
   #_w3 := "Q_Den_Run" AND "Xuat hang - Buoc 1: Di chuyen den vi tri lay";
   #_w4 := #_w3 AND NOT "P8";   // rising edge
   "P8" := #_w3;
   IF #_w4 THEN
       "Cai vi tri nhap xuat hang" := "Hien thi vi tri nhap xuat hang";
       "Xuat hang - Buoc 2: Lay hang" := TRUE;
       "Xuat hang - Buoc 1: Di chuyen den vi tri lay" := FALSE;
   END_IF;
END_REGION

REGION Network 17: Xuất hàng bước 2
   #_w1 := "Q_Den_Run" AND "Xuat hang - Buoc 2: Lay hang";
   "IEC_Timer_0_DB_7".TON(IN := #_w1, PT := T#1s);
   #_w2 := "IEC_Timer_0_DB_7".Q AND NOT "Ban nang dang moving x" AND NOT "Ban nang dang moving z";
   #_w3 := #_w2 AND NOT "P9";   // rising edge
   "P9" := #_w2;
   IF #_w3 THEN "Q_ban nang sang phai" := TRUE; END_IF;
   "IEC_Timer_0_DB_8".TON(IN := #_w1 AND "Q_ban nang sang phai", PT := T#1s);
   IF "IEC_Timer_0_DB_8".Q THEN "Q_Ban_Nang_Nang_len" := TRUE; END_IF;
   "IEC_Timer_0_DB_9".TON(IN := #_w1 AND "Q_Ban_Nang_Nang_len", PT := T#1s);
   IF "IEC_Timer_0_DB_9".Q THEN
       "TG_xuat_hang_buoc2" := TRUE;
       "Q_ban nang sang phai" := FALSE;
   END_IF;
   "IEC_Timer_0_DB_10".TON(IN := #_w1 AND "TG_xuat_hang_buoc2", PT := T#3s);
   IF "IEC_Timer_0_DB_10".Q THEN
       "Cai vi tri nhap xuat hang" := 100;
       "Xuat hang - Buoc 3: Ve vi tri home" := TRUE;
       "Xuat hang - Buoc 2: Lay hang" := FALSE;
   END_IF;
   IF NOT #_w1 THEN "TG_xuat_hang_buoc2" := FALSE; END_IF;
END_REGION

REGION Network 18: Xuất hàng bước 3
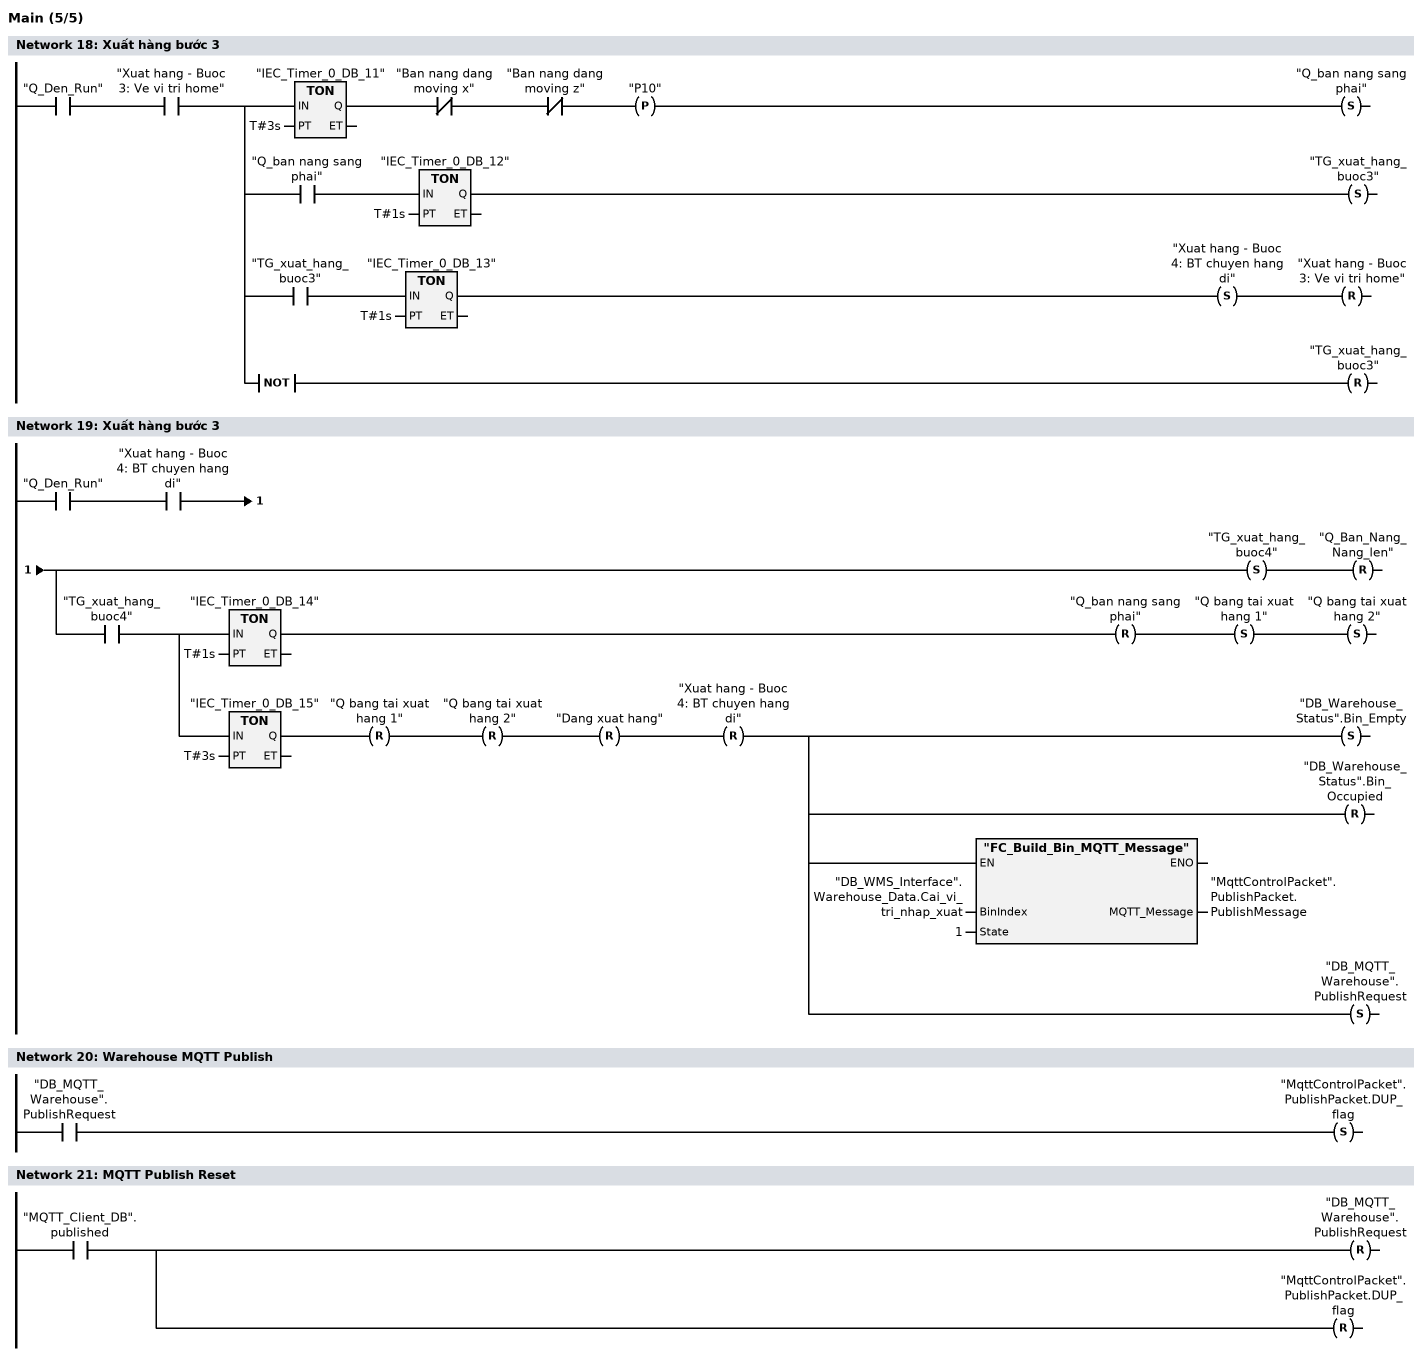
   #_w1 := "Q_Den_Run" AND "Xuat hang - Buoc 3: Ve vi tri home";
   "IEC_Timer_0_DB_11".TON(IN := #_w1, PT := T#3s);
   #_w2 := "IEC_Timer_0_DB_11".Q AND NOT "Ban nang dang moving x" AND NOT "Ban nang dang moving z";
   #_w3 := #_w2 AND NOT "P10";   // rising edge
   "P10" := #_w2;
   IF #_w3 THEN "Q_ban nang sang phai" := TRUE; END_IF;
   "IEC_Timer_0_DB_12".TON(IN := #_w1 AND "Q_ban nang sang phai", PT := T#1s);
   IF "IEC_Timer_0_DB_12".Q THEN "TG_xuat_hang_buoc3" := TRUE; END_IF;
   "IEC_Timer_0_DB_13".TON(IN := #_w1 AND "TG_xuat_hang_buoc3", PT := T#1s);
   IF "IEC_Timer_0_DB_13".Q THEN
       "Xuat hang - Buoc 4: BT chuyen hang di" := TRUE;
       "Xuat hang - Buoc 3: Ve vi tri home" := FALSE;
   END_IF;
   IF NOT #_w1 THEN "TG_xuat_hang_buoc3" := FALSE; END_IF;
END_REGION

REGION Network 19: Xuất hàng bước 3
   #_w1 := "Q_Den_Run" AND "Xuat hang - Buoc 4: BT chuyen hang di";
   IF #_w1 THEN
       "TG_xuat_hang_buoc4" := TRUE;
       "Q_Ban_Nang_Nang_len" := FALSE;
   END_IF;
   #_w2 := #_w1 AND "TG_xuat_hang_buoc4";
   "IEC_Timer_0_DB_14".TON(IN := #_w2, PT := T#1s);
   IF "IEC_Timer_0_DB_14".Q THEN
       "Q_ban nang sang phai" := FALSE;
       "Q bang tai xuat hang 1" := TRUE;
       "Q bang tai xuat hang 2" := TRUE;
   END_IF;
   "IEC_Timer_0_DB_15".TON(IN := #_w2, PT := T#3s);
   IF "IEC_Timer_0_DB_15".Q THEN
       "Q bang tai xuat hang 1" := FALSE;
       "Q bang tai xuat hang 2" := FALSE;
       "Dang xuat hang" := FALSE;
       "Xuat hang - Buoc 4: BT chuyen hang di" := FALSE;
       "DB_Warehouse_Status".Bin_Empty := TRUE;
       "DB_Warehouse_Status".Bin_Occupied := FALSE;
   END_IF;
   #_w3 := "IEC_Timer_0_DB_15".Q;
   IF #_w3 THEN
       "FC_Build_Bin_MQTT_Message"(BinIndex := "DB_WMS_Interface".Warehouse_Data.Cai_vi_tri_nhap_xuat,
                               State := 1,
                               MQTT_Message => "MqttControlPacket".PublishPacket.PublishMessage);
       "DB_MQTT_Warehouse".PublishRequest := TRUE;
   END_IF;
END_REGION

REGION Network 20: Warehouse MQTT Publish
   RUNG wire#powerrail
      Contact( "DB_MQTT_Warehouse".PublishRequest )
      S_Coil( "MqttControlPacket".PublishPacket.DUP_flag )
   END_RUNG
   // the same network as SCL:
   IF "DB_MQTT_Warehouse".PublishRequest THEN "MqttControlPacket".PublishPacket.DUP_flag := TRUE; END_IF;
END_REGION

REGION Network 21: MQTT Publish Reset
   RUNG wire#powerrail
      Contact( "MQTT_Client_DB".published )
      wire#w1
      R_Coil( "DB_MQTT_Warehouse".PublishRequest )
   END_RUNG
   RUNG wire#w1
      R_Coil( "MqttControlPacket".PublishPacket.DUP_flag )
   END_RUNG
   // the same network as SCL:
   IF "MQTT_Client_DB".published THEN
       "DB_MQTT_Warehouse".PublishRequest := FALSE;
       "MqttControlPacket".PublishPacket.DUP_flag := FALSE;
   END_IF;
END_REGION
END_ORGANIZATION_BLOCK

// folder: MqttClient

FUNCTION_BLOCK "MQTT_Client"   // FB1501, SCL
TITLE = MQTT Client
{ S7_Optimized_Access := 'TRUE' }
AUTHOR : YU_WEN_TANG
FAMILY : SLT_APC_FA
NAME : SLTAPCFA_1
VERSION : 1.0
// //============================================================================
// //Siemens Limited Taiwan 西門子台灣
// //(c)Copyright (2018) All Rights Reserved
// //----------------------------------------------------------------------------
// //Library:      MQTT client
// //Tested with:  S7-1200 FW4.2
// //Engineering:  TIA Portal V14 SP1
// //Restrictions: 
// //Requirements: SIMATIC S7-1200 FW4.0 and above
// //Functionality:
// //----------------------------------------------------------------------------
// //Change log table:
// //Version   Date        Expert in charge Changes applied
// //V1.0:     2018.04.03  SLT APC/FA YU-wen Tang 唐雨文
// //----------------------------------------------------------------------------
   VAR_INPUT
      InterfaceID : UInt;
      BrokerIP1 : Byte;
      BrokerIP2 : Byte;
      BrokerIP3 : Byte;
      BrokerIP4 : Byte;
      BrokerPort : UInt;
   END_VAR
   VAR_OUTPUT
      Busy : Bool;
      Status : Byte;
      Error : Bool;
      ErrorID : Word;
      ErrorSource : Byte;
      ReceivedTopic : Array[0..9] of String;
      ReceivedMessage : Array[0..9] of String;
   END_VAR
   VAR_IN_OUT
      Enable : Bool;
      Publish : Bool;
      Subscribe : Bool;
      Unsubscribe : Bool;
      ConnectPacket : "MqttConnectPacket";
      PublishPacket : "MqttPublishPacket";
      SubscribePacket : "MqttSubscribePacket";
      UnsubscribePacket : "MqttUnsubscribePacket";
   END_VAR
   VAR
      CONNECT : TCON_IP_v4;
      AutoPublishTimer : TON_TIME;
      TSEND_C : TSEND_C;
      TRCV : TRCV;
      TSENDATA : Array[0..499] of Byte;
      TRCVDATA : Array[0..499] of Byte;
      ConnectMsgFormat : Array[0..499] of Byte;
      PublishMsgFormat : Array[0..499] of Byte;
      SubscribeMsgFormat : Array[0..499] of Byte;
      SubscribeReqQosSetIndex : Array[0..9] of Int;
      UnsubscribeMsgFormat : Array[0..499] of Byte;
      RcvDataBuffer : Array[0..15, 0..499] of Byte;
      RcvDataNDR : Array[0..15] of Bool;
      RcvDataNDLen : Array[0..15] of UDInt;
      strg_to_chars : Array[0..253] of Char;
      p_trig : Array[0..31] of Bool;   // [7]
      WatchDogTimer : TON_TIME;
      KeepAliveTimer : TON_TIME;
      iError : Bool;
      Idle : Bool;
      TcpConnected : Bool;
      MqttConnected : Bool;
      published : Bool;
      subscribed : Bool;
      unsubscribed : Bool;
      pinged : Bool;
      disconnected : Bool;
      subscribedMsgReceived : Bool;
      watchDogEnable : Bool;
      keepAliveEnable : Bool;
      keepAliveTimerQ : Bool;
      willQoS_1 : Bool;
      willQoS_2 : Bool;
      sessionPresent : Bool;
      connectEncodedRL : Byte;
      publishEncodedRL : Byte;
      subscribeEncodedRL : Byte;
      unsubscribeEncodedRL : Byte;
      RLencodedByte : Byte;
      subscribedMsgQos : Byte;
      LengthTmp : Word;
      subscribedTopicLength_tmp : Word;
      packetIdWordTmp : Word;
      iErrorID : Word;
      ConnectReturnCode : Word;
      ConnectStep : Int;
      PublishStep : Int;
      PingReqStep : Int;
      SubscribeStep : Int;
      UnsubscribeStep : Int;
      SubscribedMsgRcvStep : Int;
      DisconnectStep : Int;
      RLencodedIndex : Int;
      subscribedMsgIndex : Int;
      subscribedTopicLength : Int;
      subscribedTopicNameIndex : Int;
      subscribedPocketIdIndex : Int;
      subscribedPayloadIndex : Int;
      RcvDataPacketType : Int;
      RcvSubscribedMsgArrayIndex : Int;
      packetID : UInt;
      strg_to_chars_cnt : UInt;
      connectRL : DInt;
      publishRL : DInt;
      subscribeRL : DInt;
      unsubscribeRL : DInt;
      connectMsgIndex : DInt;
      publishMsgIndex : DInt;
      subscribeMsgIndex : DInt;
      unsubscribeMsgIndex : DInt;
      subackDecodedRL : DInt;
      subscribedPayloadDecodedRL : DInt;
      PingReqCounter : DInt;
      PingRespCounter : DInt;
      RLmultiplier : DInt;
      subscribedPayloadLength : DInt;
      keepAliveTime : Time;
   END_VAR
   VAR_TEMP
      i : Int;
      j : Int;
   END_VAR
   // TRCV.EN_R := False;
   // TRCV.ADHOC := False;
   // TRCV.NDR := False;
   // TRCV.BUSY := False;
   // TRCV.ERROR := False;
   // TSEND_C.REQ := False;
   // TSEND_C.CONT := False;
   // TSEND_C.DONE := False;
   // TSEND_C.BUSY := False;
   // TSEND_C.ERROR := False;
   // TSEND_C.COM_RST := False;
   // KeepAliveTimer.IN := False;
   // WatchDogTimer.IN := False;
   // RcvDataNDR[15] := False;
   // RcvDataNDR[14] := False;
   // RcvDataNDR[13] := False;
   // RcvDataNDR[12] := False;
   // RcvDataNDR[11] := False;
   // RcvDataNDR[10] := False;
   // RcvDataNDR[9] := False;
   // RcvDataNDR[8] := False;
   // RcvDataNDR[7] := False;
   // RcvDataNDR[6] := False;
   // RcvDataNDR[5] := False;
   // RcvDataNDR[4] := False;
   // RcvDataNDR[3] := False;
   // RcvDataNDR[2] := False;
   // RcvDataNDR[1] := False;
   // RcvDataNDR[0] := False;
   // p_trig[31] := False;
   // p_trig[30] := False;
   // p_trig[29] := False;
   // p_trig[28] := False;
   // p_trig[27] := False;
   // p_trig[26] := False;
   // p_trig[25] := False;
   // p_trig[24] := False;
   // p_trig[23] := False;
   // p_trig[22] := False;
   // p_trig[21] := False;
   // p_trig[20] := False;
   // p_trig[19] := False;
   // p_trig[18] := False;
   // p_trig[17] := False;
   // p_trig[16] := False;
   // p_trig[15] := False;
   // p_trig[14] := False;
   // p_trig[13] := False;
   // p_trig[12] := False;
   // p_trig[11] := False;
   // p_trig[10] := False;
   // p_trig[9] := False;
   // p_trig[8] := False;
   // p_trig[7] := False;
   // p_trig[6] := False;
   // p_trig[5] := False;
   // p_trig[4] := False;
   // p_trig[3] := False;
   // p_trig[2] := False;
   // p_trig[1] := False;
   // p_trig[0] := False;
BEGIN
   //============================================================================
   //Siemens Limited Taiwan 西門子台灣
   //(c)Copyright (2018) All Rights Reserved
   //----------------------------------------------------------------------------
   //Library:      MQTT Client
   //Requirements: SIMATIC S7-1200 FW4.0 and above
   //Tested with:  S7-1200 FW4.2
   //Tested MQTT Broker: Mosquitto
   //Engineering:  TIA Portal V14 SP1
   //Restrictions: None, Free for use / modification
   //Author: Siemens Limited Taiwan DF/FA/APC, Yu-wen Tang 唐雨文
   //Date: 2018.04.03
   //----------------------------------------------------------------------------
   REGION OUC functions
       #TSEND_C(CONNECT := #CONNECT,
                CONT := True,
                DATA := #TSENDATA);
       IF (#TSEND_C.DONE AND NOT #TSEND_C.BUSY) OR #TSEND_C.ERROR THEN
           #TSEND_C.REQ := False;
       END_IF;
       #TRCV(EN_R := True,
             ID := #CONNECT.ID,
             LEN := 0,
             ADHOC := True,
             DATA := #TRCVDATA);
       IF (#TRCV.NDR AND #TRCV.RCVD_LEN > 0) AND NOT #p_trig[1] THEN
           #RcvDataPacketType := BYTE_TO_INT(SHR(IN := #TRCVDATA[0], N := 4));
           UMOVE_BLK(IN := #TRCVDATA[0],
                     COUNT := #TRCV.RCVD_LEN,
                     OUT => #RcvDataBuffer[#RcvDataPacketType, 0]);
           #RcvDataNDR[#RcvDataPacketType] := True;
           #RcvDataNDLen[#RcvDataPacketType] := #TRCV.RCVD_LEN;
       END_IF;
       #p_trig[1] := #TRCV.NDR AND #TRCV.RCVD_LEN > 0;
   END_REGION
   REGION Enable & Execute
       IF #Enable AND NOT #p_trig[0] THEN
           #CONNECT.ID := 16#0FFF;
           #CONNECT.InterfaceId := #InterfaceID;
           #CONNECT.ActiveEstablished := True;
           #CONNECT.RemoteAddress.ADDR[1] := #BrokerIP1;
           #CONNECT.RemoteAddress.ADDR[2] := #BrokerIP2;
           #CONNECT.RemoteAddress.ADDR[3] := #BrokerIP3;
           #CONNECT.RemoteAddress.ADDR[4] := #BrokerIP4;
           #CONNECT.RemotePort := #BrokerPort;
           #CONNECT.LocalPort := 0;
           #keepAliveTime := INT_TO_TIME(WORD_TO_INT(#ConnectPacket.keepAliveTime) * 1000);
           #iError := False;
           #iErrorID := 16#0000;
           #ErrorSource := 16#00;
           #TSEND_C.REQ := False;
           #Publish := False;
           #Subscribe := False;
           #Unsubscribe := False;
           #ConnectStep := 0;
           #PublishStep := 0;
           #SubscribeStep := 0;
           #UnsubscribeStep := 0;
           #PingReqStep := 0;
           #DisconnectStep := 0;
           #SubscribedMsgRcvStep := 0;
           #PingReqCounter := 0;
           #PingRespCounter := 0;
           #published := False;
           #subscribed := False;
           #unsubscribed := False;
           #pinged := False;
       END_IF;
       IF NOT #Enable AND #p_trig[0] THEN
           #published := False;
           #subscribed := False;
           #unsubscribed := False;
           #pinged := False;
           #Publish := False;
           #Subscribe := False;
           #Unsubscribe := False;
           #ConnectStep := 0;
           #PublishStep := 0;
           #SubscribeStep := 0;
           #UnsubscribeStep := 0;
           #PingReqStep := 0;
           #DisconnectStep := 1;
           #SubscribedMsgRcvStep := 0;
           #PingReqCounter := 0;
           #PingRespCounter := 0;
           #watchDogEnable := False;
           #keepAliveEnable := False;
           FOR #i := 0 TO 15 DO
               #RcvDataNDR[#i] := False;
               #RcvDataNDLen[#i] := 0;
           END_FOR;
           IF NOT #iError THEN
               #DisconnectStep := 1;
           END_IF;
       END_IF;
       #p_trig[0] := #Enable;
       #TcpConnected := #Enable AND #TSEND_C.CONT AND #TSEND_C.s_TDIAG_Status.State = 16#04;
       IF NOT #TcpConnected THEN
           #MqttConnected := False;
           #Enable := False;
       END_IF;
       IF NOT #MqttConnected THEN
           IF #Publish THEN
               #iError := True;
               #iErrorID := 16#9104;
               #ErrorSource := 16#03;
               #Publish := False;
           ELSIF #Subscribe THEN
               #iError := True;
               #iErrorID := 16#9104;
               #ErrorSource := 16#08;
               #Subscribe := False;
           ELSIF #Unsubscribe THEN
               #iError := True;
               #iErrorID := 16#9104;
               #ErrorSource := 16#0A;
               #Unsubscribe := False;
           ELSIF
               #PingReqStep > 0 THEN
               #iError := True;
               #iErrorID := 16#9104;
               #ErrorSource := 16#0C;
               #PingReqStep := 0;
           END_IF;
       END_IF;
       IF #Enable AND #TRCV.STATUS = 16#80C4 THEN
           #iError := True;
           #ErrorSource := 16#00;
           #iErrorID := #TRCV.STATUS;
           #Enable := False;
       END_IF;
       IF (#TRCV.STATUS = 16#80A1 OR #TRCV.STATUS = 16#80C6) THEN
           #iError := True;
           #ErrorSource := 16#00;
           #iErrorID := #TRCV.STATUS;
       END_IF;
       IF #iError AND NOT #p_trig[2] THEN
           #TSEND_C.REQ := False;
           #watchDogEnable := False;
           #keepAliveEnable := False;
           #Publish := False;
           #Subscribe := False;
           #Unsubscribe := False;
           IF #iErrorID > 16#9000 AND #iErrorID < 16#9100 THEN
               #DisconnectStep := 1;
           ELSE
               #Enable := False;
           END_IF;
       END_IF;
       #p_trig[2] := #iError;
       IF #TcpConnected AND #Enable AND NOT #MqttConnected AND #DisconnectStep = 0 AND NOT #p_trig[3] THEN
           #ConnectStep := 1;
       END_IF;
       #p_trig[3] := #TcpConnected AND #Enable AND NOT #MqttConnected AND #DisconnectStep = 0;
       #Idle := #ConnectStep = 0 AND #PublishStep = 0 AND #SubscribeStep = 0 AND #UnsubscribeStep = 0 AND #DisconnectStep = 0 AND #SubscribedMsgRcvStep = 0;
       IF #ConnectPacket.keepAliveTime > 16#0000 AND #ConnectPacket.keepAliveTime < 16#0002 THEN
           #ConnectPacket.keepAliveTime := 16#0002;
       END_IF;
       IF #TcpConnected AND #MqttConnected AND #Idle AND #ConnectPacket.keepAliveTime > 16#0000 THEN
           #keepAliveEnable := True;
       ELSE
           #keepAliveEnable := False;
       END_IF;
       IF #keepAliveEnable AND #keepAliveTimerQ THEN
           #PingReqStep := 1;
       END_IF;
       IF #WatchDogTimer.Q THEN
           #watchDogEnable := False;
           #iErrorID := 16#9001;
           #iError := True;
           IF #ConnectStep > 0 THEN
               #ErrorSource := 16#01;
           ELSIF #PublishStep > 0 THEN
               #ErrorSource := 16#03;
           ELSIF #SubscribeStep > 0 THEN
               #ErrorSource := 16#08;
           ELSIF #UnsubscribeStep > 0 THEN
               #ErrorSource := 16#0A;
           ELSIF #PingReqStep > 0 THEN
               #ErrorSource := 16#0C;
           ELSIF #DisconnectStep > 0 THEN
               #ErrorSource := 16#0E;
           ELSIF #SubscribedMsgRcvStep > 0 THEN
               #ErrorSource := 16#0F;
           END_IF;
       END_IF;
   END_REGION ;
   REGION CONNECT
       CASE #ConnectStep OF
           0:
               ;
           1:
               #PingReqStep := 0;
               #iError := False;
               #iErrorID := 16#0000;
               #ErrorSource := 16#00;
               #ConnectStep := 2;
           2:
               IF #ConnectPacket.willFlag THEN
                   CASE #ConnectPacket.willQoS_level OF
                       0:
                           #willQoS_1 := False;
                           #willQoS_2 := False;
                       1:
                           #willQoS_1 := True;
                           #willQoS_2 := False;
                       2:
                           #willQoS_1 := False;
                           #willQoS_2 := True;
                       ELSE
                           #iError := True;
                           #iErrorID := 16#9100;
                           #ErrorSource := 16#01;
                           #ConnectStep := 13;
                   END_CASE;
               ELSE
                   #willQoS_1 := False;
                   #willQoS_2 := False;
                   #ConnectPacket.willRetain := False;
               END_IF;
               #ConnectStep := 3;
           3:
               #connectRL := 12;
               #ConnectPacket.cleanSession := True;
               IF #ConnectPacket.clientIdentifier = '' OR LEN(#ConnectPacket.clientIdentifier) > 23 THEN
                   #iError := True;
                   #iErrorID := 16#9107;
                   #ErrorSource := 16#01;
                   #ConnectStep := 13;
               END_IF;
               #connectRL := #connectRL + LEN(#ConnectPacket.clientIdentifier);
               IF #ConnectPacket.willFlag THEN
                   IF #ConnectPacket.willTopic = '' THEN
                       #iError := True;
                       #iErrorID := 16#9108;
                       #ErrorSource := 16#01;
                       #ConnectStep := 13;
                   END_IF;
                   #connectRL := #connectRL + 2 + LEN(#ConnectPacket.willTopic) + 2 + LEN(#ConnectPacket.willMessage);
               END_IF;
               IF #ConnectPacket.userNameFlag THEN
                   #connectRL := #connectRL + LEN(#ConnectPacket.userName);
                   #connectRL := #connectRL + 2;
               ELSE
                   #ConnectPacket.passwordFlag := False;
               END_IF;
               IF #ConnectPacket.passwordFlag THEN
                   #connectRL := #connectRL + LEN(#ConnectPacket.password);
                   #connectRL := #connectRL + 2;
               END_IF;
               #ConnectStep := 4;
           4:
               #ConnectMsgFormat[0] := 16#10;
               #ConnectStep := 5;
           5:
               #connectMsgIndex := 1;
               REPEAT
                   #connectEncodedRL := DINT_TO_BYTE(#connectRL MOD 128);
                   #connectRL := #connectRL / 128;
                   IF #connectRL > 0 THEN
                       #connectEncodedRL := #connectEncodedRL OR 128;
                       #ConnectMsgFormat[#connectMsgIndex] := #connectEncodedRL;
                       #connectMsgIndex := #connectMsgIndex + 1;
                   ELSE
                       #ConnectMsgFormat[#connectMsgIndex] := #connectEncodedRL;
                   END_IF;
               UNTIL #connectRL <= 0 END_REPEAT;
               #ConnectStep := 6;
           6:
               #connectMsgIndex := #connectMsgIndex + 1;
               #ConnectMsgFormat[#connectMsgIndex] := 0;
               #connectMsgIndex := #connectMsgIndex + 1;
               #ConnectMsgFormat[#connectMsgIndex] := 4;
               #connectMsgIndex := #connectMsgIndex + 1;
               #ConnectMsgFormat[#connectMsgIndex] := CHAR_TO_BYTE('M');
               #connectMsgIndex := #connectMsgIndex + 1;
               #ConnectMsgFormat[#connectMsgIndex] := CHAR_TO_BYTE('Q');
               #connectMsgIndex := #connectMsgIndex + 1;
               #ConnectMsgFormat[#connectMsgIndex] := CHAR_TO_BYTE('T');
               #connectMsgIndex := #connectMsgIndex + 1;
               #ConnectMsgFormat[#connectMsgIndex] := CHAR_TO_BYTE('T');
               #connectMsgIndex := #connectMsgIndex + 1;
               #ConnectMsgFormat[#connectMsgIndex] := 16#04;
               #connectMsgIndex := #connectMsgIndex + 1;
               #ConnectMsgFormat[#connectMsgIndex].%X0 := False;
               #ConnectMsgFormat[#connectMsgIndex].%X1 := #ConnectPacket.cleanSession;
               #ConnectMsgFormat[#connectMsgIndex].%X2 := #ConnectPacket.willFlag;
               #ConnectMsgFormat[#connectMsgIndex].%X3 := #willQoS_1;
               #ConnectMsgFormat[#connectMsgIndex].%X4 := #willQoS_2;
               #ConnectMsgFormat[#connectMsgIndex].%X5 := #ConnectPacket.willRetain;
               IF NOT #ConnectMsgFormat[#connectMsgIndex].%X7 THEN
                   #ConnectPacket.passwordFlag := False;
               END_IF;
               #ConnectMsgFormat[#connectMsgIndex].%X6 := #ConnectPacket.passwordFlag;
               #ConnectMsgFormat[#connectMsgIndex].%X7 := #ConnectPacket.userNameFlag;
               #connectMsgIndex := #connectMsgIndex + 1;
               #ConnectMsgFormat[#connectMsgIndex] := #ConnectPacket.keepAliveTime.%B1;
               #connectMsgIndex := #connectMsgIndex + 1;
               #ConnectMsgFormat[#connectMsgIndex] := #ConnectPacket.keepAliveTime.%B0;
               #connectMsgIndex := #connectMsgIndex + 1;
               #LengthTmp := INT_TO_WORD(LEN(#ConnectPacket.clientIdentifier));
               #ConnectMsgFormat[#connectMsgIndex] := #LengthTmp.%B1;
               #connectMsgIndex := #connectMsgIndex + 1;
               #ConnectMsgFormat[#connectMsgIndex] := #LengthTmp.%B0;
               Strg_TO_Chars(Strg := #ConnectPacket.clientIdentifier,
                             pChars := 0,
                             Cnt => #strg_to_chars_cnt,
                             Chars := #strg_to_chars);
               FOR #i := 0 TO UINT_TO_INT(#strg_to_chars_cnt) - 1 DO
                   #connectMsgIndex := #connectMsgIndex + 1;
                   #ConnectMsgFormat[#connectMsgIndex] := CHAR_TO_BYTE(#strg_to_chars[#i]);
               END_FOR;
               IF #ConnectPacket.willFlag THEN
                   #LengthTmp := INT_TO_WORD(LEN(#ConnectPacket.willTopic));
                   #connectMsgIndex := #connectMsgIndex + 1;
                   #ConnectMsgFormat[#connectMsgIndex] := #LengthTmp.%B1;
                   #connectMsgIndex := #connectMsgIndex + 1;
                   #ConnectMsgFormat[#connectMsgIndex] := #LengthTmp.%B0;
                   Strg_TO_Chars(Strg := #ConnectPacket.willTopic,
                                 pChars := 0,
                                 Cnt => #strg_to_chars_cnt,
                                 Chars := #strg_to_chars);
                   FOR #i := 0 TO UINT_TO_INT(#strg_to_chars_cnt) - 1 DO
                       #connectMsgIndex := #connectMsgIndex + 1;
                       #ConnectMsgFormat[#connectMsgIndex] := CHAR_TO_BYTE(#strg_to_chars[#i]);
                   END_FOR;
                   #LengthTmp := INT_TO_WORD(LEN(#ConnectPacket.willMessage));
                   #connectMsgIndex := #connectMsgIndex + 1;
                   #ConnectMsgFormat[#connectMsgIndex] := #LengthTmp.%B1;
                   #connectMsgIndex := #connectMsgIndex + 1;
                   #ConnectMsgFormat[#connectMsgIndex] := #LengthTmp.%B0;
                   Strg_TO_Chars(Strg := #ConnectPacket.willMessage,
                                 pChars := 0,
                                 Cnt => #strg_to_chars_cnt,
                                 Chars := #strg_to_chars);
                   FOR #i := 0 TO UINT_TO_INT(#strg_to_chars_cnt) - 1 DO
                       #connectMsgIndex := #connectMsgIndex + 1;
                       #ConnectMsgFormat[#connectMsgIndex] := CHAR_TO_BYTE(#strg_to_chars[#i]);
                   END_FOR;
               END_IF;
               IF #ConnectPacket.userNameFlag THEN
                   #LengthTmp := INT_TO_WORD(LEN(#ConnectPacket.userName));
                   #connectMsgIndex := #connectMsgIndex + 1;
                   #ConnectMsgFormat[#connectMsgIndex] := #LengthTmp.%B1;
                   #connectMsgIndex := #connectMsgIndex + 1;
                   #ConnectMsgFormat[#connectMsgIndex] := #LengthTmp.%B0;
                   Strg_TO_Chars(Strg := #ConnectPacket.userName,
                                 pChars := 0,
                                 Cnt => #strg_to_chars_cnt,
                                 Chars := #strg_to_chars);
                   FOR #i := 0 TO UINT_TO_INT(#strg_to_chars_cnt) - 1 DO
                       #connectMsgIndex := #connectMsgIndex + 1;
                       #ConnectMsgFormat[#connectMsgIndex] := CHAR_TO_BYTE(#strg_to_chars[#i]);
                   END_FOR;
               END_IF;
               IF #ConnectPacket.passwordFlag THEN
                   #LengthTmp := INT_TO_WORD(LEN(#ConnectPacket.password));
                   #connectMsgIndex := #connectMsgIndex + 1;
                   #ConnectMsgFormat[#connectMsgIndex] := #LengthTmp.%B1;
                   #connectMsgIndex := #connectMsgIndex + 1;
                   #ConnectMsgFormat[#connectMsgIndex] := #LengthTmp.%B0;
                   Strg_TO_Chars(Strg := #ConnectPacket.password,
                                 pChars := 0,
                                 Cnt => #strg_to_chars_cnt,
                                 Chars := #strg_to_chars);
                   FOR #i := 0 TO UINT_TO_INT(#strg_to_chars_cnt) - 1 DO
                       #connectMsgIndex := #connectMsgIndex + 1;
                       #ConnectMsgFormat[#connectMsgIndex] := CHAR_TO_BYTE(#strg_to_chars[#i]);
                   END_FOR;
               END_IF;
               #ConnectStep := 7;
           7:
               UMOVE_BLK(IN := #ConnectMsgFormat[0],
                         COUNT := DINT_TO_UINT(#connectMsgIndex + 1),
                         OUT => #TSENDATA[0]);
               #ConnectStep := 8;
           8:
               UFILL_BLK(IN := 16#00,
                         COUNT := 255,
                         OUT => #RcvDataBuffer[2, 0]);
               #ConnectStep := 9;
           9:
               #TSEND_C.LEN := DINT_TO_UINT(#connectMsgIndex + 1);
               #RcvDataNDR[2] := False;
               #RcvDataNDLen[2] := 0;
               #TSEND_C.REQ := True;
               #ConnectStep := 10;
           10:
               #watchDogEnable := True;
               IF #TSEND_C.DONE AND NOT #TSEND_C.BUSY THEN
                   #ConnectStep := 11;
               END_IF;
           11:
               IF #RcvDataNDR[2] AND #RcvDataNDLen[2] > 0 THEN
                   #watchDogEnable := False;
                   #sessionPresent := #RcvDataBuffer[2, 2].%X0;
                   #ConnectReturnCode := #RcvDataBuffer[2, 3];
                   IF #RcvDataBuffer[2, 0] = 16#20 AND #RcvDataBuffer[2, 1] = 16#02 AND #RcvDataBuffer[2, 2] < 2 THEN
                       #ConnectStep := 12;
                   ELSE
                       #iError := True;
                       #iErrorID := 16#9003;
                       #ErrorSource := 16#02;
                       #ConnectStep := 13;
                   END_IF;
                   IF #ConnectReturnCode <> 16#00 THEN
                       #iError := True;
                       #iErrorID := 16#9004;
                       #ErrorSource := 16#02;
                       #ConnectStep := 13;
                   END_IF;
               END_IF;
           12:
               #MqttConnected := True;
               #ConnectStep := 13;
           13:
               #RcvDataNDR[2] := False;
               #RcvDataNDLen[2] := 0;
               #ConnectStep := 0;
               #watchDogEnable := False;
       END_CASE;
   END_REGION ;
   REGION PUBLISH
       IF #MqttConnected AND #Publish AND #Idle AND NOT #p_trig[4] THEN
           #PublishStep := 1;
       END_IF;
       #p_trig[4] := #MqttConnected AND #Publish AND #Idle;
       CASE #PublishStep OF
           0:
               ;
           1:
               #published := False;
               #subscribed := False;
               #unsubscribed := False;
               #pinged := False;
               #disconnected := False;
               #subscribedMsgReceived := False;
               IF #PublishPacket.PublishTopic = '' THEN
                   #iError := True;
                   #iErrorID := 16#9101;
                   #ErrorSource := 16#03;
                   #PublishStep := 40;
               ELSE
                   #PingReqStep := 0;
                   #iError := False;
                   #iErrorID := 16#0000;
                   #ErrorSource := 16#00;
                   #PublishStep := 2;
               END_IF;
           2:
               #publishRL := 2;
               #publishRL := #publishRL + LEN(#PublishPacket.PublishTopic);
               #publishRL := #publishRL + LEN(#PublishPacket.PublishMessage);
               #PublishStep := 3;
           3:
               #PublishMsgFormat[0] := 16#30;
               CASE #PublishPacket.QoS_level OF
                   0:
                       #PublishMsgFormat[0].%X1 := False;
                       #PublishMsgFormat[0].%X2 := False;
                       #PublishPacket.DUP_flag := False;
                   1:
                       #PublishMsgFormat[0].%X1 := True;
                       #PublishMsgFormat[0].%X2 := False;
                       #publishRL := #publishRL + 2;
                   2:
                       #PublishMsgFormat[0].%X1 := False;
                       #PublishMsgFormat[0].%X2 := True;
                       #publishRL := #publishRL + 2;
                   ELSE
                       #iError := True;
                       #iErrorID := 16#9102;
                       #ErrorSource := 16#03;
                       #PublishStep := 40;
               END_CASE;
               #PublishMsgFormat[0].%X0 := #PublishPacket.Retain;
               #PublishMsgFormat[0].%X3 := #PublishPacket.DUP_flag;
               #PublishStep := 4;
           4:
               #publishMsgIndex := 1;
               REPEAT
                   #publishEncodedRL := DINT_TO_BYTE(#publishRL MOD 128);
                   #publishRL := #publishRL / 128;
                   IF #publishRL > 0 THEN
                       #publishEncodedRL := #publishEncodedRL OR 128;
                       #PublishMsgFormat[#publishMsgIndex] := #publishEncodedRL;
                       #publishMsgIndex := #publishMsgIndex + 1;
                   ELSE
                       #PublishMsgFormat[#publishMsgIndex] := #publishEncodedRL;
                   END_IF;
               UNTIL #publishRL <= 0 END_REPEAT;
               #PublishStep := 5;
           5:
               #LengthTmp := INT_TO_WORD(LEN(#PublishPacket.PublishTopic));
               #publishMsgIndex := #publishMsgIndex + 1;
               #PublishMsgFormat[#publishMsgIndex] := #LengthTmp.%B1;
               #publishMsgIndex := #publishMsgIndex + 1;
               #PublishMsgFormat[#publishMsgIndex] := #LengthTmp.%B0;
               Strg_TO_Chars(Strg := #PublishPacket.PublishTopic,
                             pChars := 0,
                             Cnt => #strg_to_chars_cnt,
                             Chars := #strg_to_chars);
               FOR #i := 0 TO UINT_TO_INT(#strg_to_chars_cnt) - 1 DO
                   #publishMsgIndex := #publishMsgIndex + 1;
                   #PublishMsgFormat[#publishMsgIndex] := CHAR_TO_BYTE(#strg_to_chars[#i]);
               END_FOR;
               #packetID := #packetID + 1;
               IF #packetID > 65535 THEN
                   #packetID := 1;
               END_IF;
               IF #PublishPacket.QoS_level > 0 THEN
                   #publishMsgIndex := #publishMsgIndex + 1;
                   #packetIdWordTmp := UINT_TO_WORD(#packetID);
                   #PublishMsgFormat[#publishMsgIndex] := #packetIdWordTmp.%B1;
                   #publishMsgIndex := #publishMsgIndex + 1;
                   #PublishMsgFormat[#publishMsgIndex] := #packetIdWordTmp.%B0;
               END_IF;
               Strg_TO_Chars(Strg := #PublishPacket.PublishMessage,
                             pChars := 0,
                             Cnt => #strg_to_chars_cnt,
                             Chars := #strg_to_chars);
               FOR #i := 0 TO UINT_TO_INT(#strg_to_chars_cnt) - 1 DO
                   #publishMsgIndex := #publishMsgIndex + 1;
                   #PublishMsgFormat[#publishMsgIndex] := CHAR_TO_BYTE(#strg_to_chars[#i]);
               END_FOR;
               #PublishStep := 6;
           6:
               UMOVE_BLK(IN := #PublishMsgFormat[0],
                         COUNT := DINT_TO_UINT(#publishMsgIndex + 1),
                         OUT => #TSENDATA[0]);
               #PublishStep := 7;
           7:
               FOR #i := 4 TO 7 DO
                   UFILL_BLK(IN := 16#00,
                             COUNT := 255,
                             OUT => #RcvDataBuffer[#i, 0]);
                   #RcvDataNDR[#i] := False;
                   #RcvDataNDLen[#i] := 0;
               END_FOR;
               #PublishStep := 8;
           8:
               #TSEND_C.LEN := DINT_TO_UINT(#publishMsgIndex + 1);
               #TSEND_C.REQ := True;
               #PublishStep := 9;
           9:
               #watchDogEnable := True;
               IF #TSEND_C.DONE AND NOT #TSEND_C.BUSY THEN
                   #PublishStep := 10;
               END_IF;
           10:
               IF #PublishPacket.QoS_level = 0 THEN
                   #PublishStep := 40;
               ELSIF #RcvDataNDR[4] OR #RcvDataNDR[5] OR #RcvDataNDR[6] OR #RcvDataNDR[7] THEN
                   #watchDogEnable := False;
                   CASE #PublishPacket.QoS_level OF
                       1:
                           #PublishStep := 30;
                       2:
                           #PublishStep := 20;
                   END_CASE;
               END_IF;
           20:
               IF #RcvDataBuffer[5, 0] = 16#50 AND #RcvDataBuffer[5, 1] = 16#02 AND #RcvDataBuffer[5, 2] = #packetIdWordTmp.%B1 AND #RcvDataBuffer[5, 3] = #packetIdWordTmp.%B0 THEN
                   #PublishStep := 21;
               ELSE
                   #iError := True;
                   #iErrorID := 16#9011;
                   #ErrorSource := 16#05;
                   #PublishStep := 40;
               END_IF;
           21:
               #TSENDATA[0] := 16#62;
               #TSENDATA[1] := 16#02;
               #TSENDATA[2] := #packetIdWordTmp.%B1;
               #TSENDATA[3] := #packetIdWordTmp.%B0;
               UFILL_BLK(IN := 16#00,
                         COUNT := 255,
                         OUT => #RcvDataBuffer[7, 0]);
               #PublishStep := 22;
           22:
               #TSEND_C.LEN := 4;
               #TSEND_C.REQ := True;
               #PublishStep := 23;
           23:
               #watchDogEnable := True;
               IF #TSEND_C.DONE AND NOT #TSEND_C.BUSY THEN
                   #PublishStep := 24;
               END_IF;
           24:
               IF #RcvDataNDR[7] THEN
                   #watchDogEnable := False;
                   IF #RcvDataBuffer[7, 0] = 16#70 AND #RcvDataBuffer[7, 1] = 16#02 AND #RcvDataBuffer[7, 2] = #packetIdWordTmp.%B1 AND #RcvDataBuffer[7, 3] = #packetIdWordTmp.%B0
                   THEN
                       #PublishStep := 40;
                   ELSE
                       #iError := True;
                       #iErrorID := 16#9012;
                       #ErrorSource := 16#07;
                       #PublishStep := 40;
                   END_IF;
               END_IF;
           30:
               IF #RcvDataBuffer[4, 0] = 16#40 AND #RcvDataBuffer[4, 1] = 16#02 AND #RcvDataBuffer[4, 2] = #packetIdWordTmp.%B1 AND #RcvDataBuffer[4, 3] = #packetIdWordTmp.%B0 THEN
                   #watchDogEnable := False;
                   #PublishStep := 40;
               ELSE
                   #iError := True;
                   #iErrorID := 16#9013;
                   #ErrorSource := 16#04;
                   #PublishStep := 40;
               END_IF;
               #PublishStep := 40;
           40:
               FOR #i := 4 TO 7 DO
                   #RcvDataNDR[#i] := False;
                   #RcvDataNDLen[#i] := 0;
               END_FOR;
               #PublishStep := 0;
               #Publish := False;
               #published := True;
               #watchDogEnable := False;
       END_CASE;
   END_REGION ;
   REGION SUBSCRIBE
       IF #MqttConnected AND #Subscribe AND #Idle AND NOT #p_trig[6] THEN
           #SubscribeStep := 1;
       END_IF;
       #p_trig[6] := #MqttConnected AND #Subscribe AND #Idle;
       CASE #SubscribeStep OF
           0:
               ;
           1:
               #published := False;
               #subscribed := False;
               #unsubscribed := False;
               #pinged := False;
               #disconnected := False;
               #subscribedMsgReceived := False;
               #PingReqStep := 0;
               #iError := False;
               #iErrorID := 16#0000;
               #ErrorSource := 16#00;
               #SubscribeStep := 2;
           2:
               #subscribeRL := 2;
               #j := 0;
               FOR #i := 0 TO 9 DO
                   IF #SubscribePacket.TopicFilter[#i] <> '' THEN
                       #SubscribeReqQosSetIndex[#j] := #i;
                       #j := #j + 1;
                       #subscribeRL := #subscribeRL + 2;
                       #subscribeRL := #subscribeRL + LEN(#SubscribePacket.TopicFilter[#i]) + 1;
                   END_IF;
               END_FOR;
               IF #j = 0 THEN
                   #iError := True;
                   #iErrorID := 16#9103;
                   #ErrorSource := 16#08;
                   #SubscribeStep := 15;
               ELSE
                   #SubscribeStep := 3;
               END_IF;
           3:
               #SubscribeMsgFormat[0] := 16#82;
               #SubscribeStep := 4;
           4:
               #subscribeMsgIndex := 1;
               REPEAT
                   #subscribeEncodedRL := DINT_TO_BYTE(#subscribeRL MOD 128);
                   #subscribeRL := #subscribeRL / 128;
                   IF #subscribeRL > 0 THEN
                       #subscribeEncodedRL := #subscribeEncodedRL OR 128;
                       #SubscribeMsgFormat[#subscribeMsgIndex] := #subscribeEncodedRL;
                       #subscribeMsgIndex := #subscribeMsgIndex + 1;
                   ELSE
                       #SubscribeMsgFormat[#subscribeMsgIndex] := #subscribeEncodedRL;
                   END_IF;
               UNTIL #subscribeRL <= 0 END_REPEAT;
               #SubscribeStep := 5;
           5:
               #packetID := #packetID + 1;
               IF #packetID > 65535 THEN
                   #packetID := 1;
               END_IF;
               #subscribeMsgIndex := #subscribeMsgIndex + 1;
               #packetIdWordTmp := UINT_TO_WORD(#packetID);
               #SubscribeMsgFormat[#subscribeMsgIndex] := #packetIdWordTmp.%B1;
               #subscribeMsgIndex := #subscribeMsgIndex + 1;
               #SubscribeMsgFormat[#subscribeMsgIndex] := #packetIdWordTmp.%B0;
               #SubscribeStep := 6;
           6:
               FOR #i := 0 TO 9 DO
                   IF #SubscribePacket.TopicFilter[#i] <> '' THEN
                       #subscribeMsgIndex := #subscribeMsgIndex + 1;
                       #LengthTmp := DINT_TO_WORD(LEN(#SubscribePacket.TopicFilter[#i]));
                       #SubscribeMsgFormat[#subscribeMsgIndex] := #LengthTmp.%B1;
                       #subscribeMsgIndex := #subscribeMsgIndex + 1;
                       #SubscribeMsgFormat[#subscribeMsgIndex] := #LengthTmp.%B0;
                       Strg_TO_Chars(Strg := #SubscribePacket.TopicFilter[#i],
                                     pChars := 0,
                                     Cnt => #strg_to_chars_cnt,
                                     Chars := #strg_to_chars);
                       FOR #j := 0 TO UINT_TO_INT(#strg_to_chars_cnt) - 1 DO
                           #subscribeMsgIndex := #subscribeMsgIndex + 1;
                           #SubscribeMsgFormat[#subscribeMsgIndex] := CHAR_TO_BYTE(#strg_to_chars[#j]);
                       END_FOR;
                       IF #SubscribePacket.RequestedQoS[#i] > 2 THEN
                           #iError := True;
                           #iErrorID := 16#9105;
                           #ErrorSource := 16#08;
                           #SubscribeStep := 15;
                       END_IF;
                       #subscribeMsgIndex := #subscribeMsgIndex + 1;
                       #SubscribeMsgFormat[#subscribeMsgIndex] := #SubscribePacket.RequestedQoS[#i];
                   END_IF;
               END_FOR;
               #SubscribeStep := 7;
           7:
               UMOVE_BLK(IN := #SubscribeMsgFormat[0],
                         COUNT := DINT_TO_UINT(#subscribeMsgIndex + 1),
                         OUT => #TSENDATA[0]);
               #SubscribeStep := 8;
           8:
               UFILL_BLK(IN := 16#00,
                         COUNT := 255,
                         OUT => #RcvDataBuffer[9, 0]);
               #SubscribeStep := 9;
           9:
               #TSEND_C.LEN := DINT_TO_UINT(#subscribeMsgIndex + 1);
               #RcvDataNDR[9] := False;
               #RcvDataNDLen[9] := 0;
               #TSEND_C.REQ := True;
               #SubscribeStep := 10;
           10:
               #watchDogEnable := True;
               IF #TSEND_C.DONE AND NOT #TSEND_C.BUSY THEN
                   #SubscribeStep := 11;
               END_IF;
           11:
               IF #RcvDataNDR[9] AND #RcvDataNDLen[9] > 0 THEN
                   #watchDogEnable := False;
                   IF #RcvDataBuffer[9, 0] = 16#90 THEN
                       #SubscribeStep := 12;
                   ELSE
                       #iError := True;
                       #iErrorID := 16#9021;
                       #ErrorSource := 16#09;
                       #SubscribeStep := 15;
                   END_IF;
               END_IF;
           12:
               #RLmultiplier := 1;
               #subackDecodedRL := 0;
               #RLencodedIndex := 1;
               REPEAT
                   #RLencodedByte := #RcvDataBuffer[9, #RLencodedIndex];
                   #subackDecodedRL := #subackDecodedRL + (BYTE_TO_DINT(#RLencodedByte AND 127) * #RLmultiplier);
                   #RLmultiplier := #RLmultiplier * 128;
                   #RLencodedIndex := #RLencodedIndex + 1;
                   IF #RLmultiplier > 128 ** 3 THEN
                       #iError := True;
                       #iErrorID := 16#9022;
                       #ErrorSource := 16#09;
                       #SubscribeStep := 15;
                   END_IF;
               UNTIL (#RLencodedByte AND 128) = 0 END_REPEAT;
               IF NOT #iError THEN
                   #SubscribeStep := 13;
               END_IF;
           13:
               IF #RcvDataBuffer[9, 2] = #packetIdWordTmp.%B1 AND #RcvDataBuffer[9, 3] = #packetIdWordTmp.%B0 THEN
                   #SubscribeStep := 14;
               ELSE
                   #iError := True;
                   #iErrorID := 16#9023;
                   #ErrorSource := 16#09;
                   #SubscribeStep := 15;
               END_IF;
           14:
               #j := 0;
               FOR #i := 4 TO (3 + DINT_TO_INT(#subackDecodedRL) - 2) DO
                   IF NOT (#RcvDataBuffer[9, #i] = #SubscribePacket.RequestedQoS[#SubscribeReqQosSetIndex[#j]]) THEN
                       #iError := True;
                       #iErrorID := 16#9024;
                       #ErrorSource := 16#09;
                       #SubscribeStep := 15;
                   END_IF;
                   #j := #j + 1;
               END_FOR;
               IF NOT #iError THEN
                   #SubscribeStep := 15;
               END_IF;
           15:
               #RcvDataNDR[9] := False;
               #RcvDataNDLen[9] := 0;
               #SubscribeStep := 0;
               #Subscribe := False;
               #subscribed := True;
               #watchDogEnable := False;
       END_CASE;
   END_REGION ;
   REGION UNSUBSCRIBE
       IF #MqttConnected AND #Unsubscribe AND #Idle AND NOT #p_trig[7] THEN
           #UnsubscribeStep := 1;
       END_IF;
       #p_trig[7] := #MqttConnected AND #Unsubscribe AND #Idle;
       CASE #UnsubscribeStep OF
           0:
               ;
           1:
               #published := False;
               #subscribed := False;
               #unsubscribed := False;
               #pinged := False;
               #disconnected := False;
               #subscribedMsgReceived := False;
               #PingReqStep := 0;
               #iError := False;
               #iErrorID := 16#0000;
               #ErrorSource := 16#00;
               #UnsubscribeStep := 2;
           2:
               #unsubscribeRL := 2;
               #j := 0;
               FOR #i := 0 TO 9 DO
                   IF #UnsubscribePacket.TopicFilter[#i] <> '' THEN
                       #unsubscribeRL := #unsubscribeRL + 2;
                       #unsubscribeRL := #unsubscribeRL + LEN(#UnsubscribePacket.TopicFilter[#i]);
                       #j := #j + 1;
                   END_IF;
               END_FOR;
               IF #j = 0 THEN
                   #iError := True;
                   #iErrorID := 16#9106;
                   #ErrorSource := 16#0B;
                   #UnsubscribeStep := 13;
               ELSE
                   #UnsubscribeStep := 3;
               END_IF;
           3:
               #UnsubscribeMsgFormat[0] := 16#A2;
               #UnsubscribeStep := 4;
           4:
               #unsubscribeMsgIndex := 1;
               REPEAT
                   #unsubscribeEncodedRL := DINT_TO_BYTE(#unsubscribeRL MOD 128);
                   #unsubscribeRL := #subscribeRL / 128;
                   IF #subscribeRL > 0 THEN
                       #unsubscribeEncodedRL := #unsubscribeEncodedRL OR 128;
                       #UnsubscribeMsgFormat[#unsubscribeMsgIndex] := #unsubscribeEncodedRL;
                       #unsubscribeMsgIndex := #unsubscribeMsgIndex + 1;
                   ELSE
                       #UnsubscribeMsgFormat[#unsubscribeMsgIndex] := #unsubscribeEncodedRL;
                   END_IF;
               UNTIL #unsubscribeRL <= 0 END_REPEAT;
               #UnsubscribeStep := 5;
           5:
               #packetID := #packetID + 1;
               IF #packetID > 65535 THEN
                   #packetID := 1;
               END_IF;
               #unsubscribeMsgIndex := #unsubscribeMsgIndex + 1;
               #packetIdWordTmp := UINT_TO_WORD(#packetID);
               #UnsubscribeMsgFormat[#unsubscribeMsgIndex] := #packetIdWordTmp.%B1;
               #unsubscribeMsgIndex := #unsubscribeMsgIndex + 1;
               #UnsubscribeMsgFormat[#unsubscribeMsgIndex] := #packetIdWordTmp.%B0;
               #UnsubscribeStep := 6;
           6:
               FOR #i := 0 TO 9 DO
                   IF #UnsubscribePacket.TopicFilter[#i] <> '' THEN
                       #unsubscribeMsgIndex := #unsubscribeMsgIndex + 1;
                       #LengthTmp := DINT_TO_WORD(LEN(#UnsubscribePacket.TopicFilter[#i]));
                       #UnsubscribeMsgFormat[#unsubscribeMsgIndex] := #LengthTmp.%B1;
                       #unsubscribeMsgIndex := #unsubscribeMsgIndex + 1;
                       #UnsubscribeMsgFormat[#unsubscribeMsgIndex] := #LengthTmp.%B0;
                       Strg_TO_Chars(Strg := #UnsubscribePacket.TopicFilter[#i],
                                     pChars := 0,
                                     Cnt => #strg_to_chars_cnt,
                                     Chars := #strg_to_chars);
                       FOR #j := 0 TO UINT_TO_INT(#strg_to_chars_cnt) - 1 DO
                           #unsubscribeMsgIndex := #unsubscribeMsgIndex + 1;
                           #UnsubscribeMsgFormat[#unsubscribeMsgIndex] := CHAR_TO_BYTE(#strg_to_chars[#j]);
                       END_FOR;
                   END_IF;
               END_FOR;
               #UnsubscribeStep := 7;
           7:
               UMOVE_BLK(IN := #UnsubscribeMsgFormat[0],
                         COUNT := DINT_TO_UINT(#unsubscribeMsgIndex + 1),
                         OUT => #TSENDATA[0]);
               #UnsubscribeStep := 8;
           8:
               UFILL_BLK(IN := 16#00,
                         COUNT := 255,
                         OUT => #RcvDataBuffer[11, 0]);
               #UnsubscribeStep := 9;
           9:
               #TSEND_C.LEN := DINT_TO_UINT(#unsubscribeMsgIndex + 1);
               #RcvDataNDR[11] := False;
               #RcvDataNDLen[11] := 0;
               #TSEND_C.REQ := True;
               #UnsubscribeStep := 10;
           10:
               #watchDogEnable := True;
               IF #TSEND_C.DONE AND NOT #TSEND_C.BUSY THEN
                   #UnsubscribeStep := 11;
               END_IF;
           11:
               IF #RcvDataNDR[11] AND #RcvDataNDLen[11] > 0 THEN
                   #watchDogEnable := False;
                   IF #RcvDataBuffer[11, 0] = 16#B0 AND #RcvDataBuffer[11, 1] = 16#02 THEN
                       #UnsubscribeStep := 12;
                   ELSE
                       #iError := True;
                       #iErrorID := 16#9030;
                       #ErrorSource := 16#11;
                       #UnsubscribeStep := 13;
                   END_IF;
               END_IF;
           12:
               IF NOT (#RcvDataBuffer[11, 2] = #packetIdWordTmp.%B1 AND #RcvDataBuffer[11, 3] = #packetIdWordTmp.%B0) THEN
                   #iError := True;
                   #iErrorID := 16#9025;
                   #ErrorSource := 16#11;
               END_IF;
               #UnsubscribeStep := 13;
           13:
               #RcvDataNDR[11] := False;
               #RcvDataNDLen[11] := 0;
               #UnsubscribeStep := 0;
               #Unsubscribe := False;
               #unsubscribed := True;
               #watchDogEnable := False;
       END_CASE;
   END_REGION ;
   REGION PINGREQ
       CASE #PingReqStep OF
           0:
               ;
           1:
               #published := False;
               #subscribed := False;
               #unsubscribed := False;
               #pinged := False;
               #disconnected := False;
               #subscribedMsgReceived := False;
               #iError := False;
               #iErrorID := 16#0000;
               #ErrorSource := 16#00;
               #PingReqStep := 2;
           2:
               #TSENDATA[0] := 16#C0;
               #TSENDATA[1] := 16#00;
               #PingReqStep := 3;
           3:
               UFILL_BLK(IN := 16#00,
                         COUNT := 500,
                         OUT => #RcvDataBuffer[13, 0]);
               #RcvDataNDR[13] := False;
               #RcvDataNDLen[13] := 0;
               #TSEND_C.LEN := 2;
               #TSEND_C.REQ := True;
               #PingReqCounter := #PingReqCounter + 1;
               #PingReqStep := 4;
           4:
               #watchDogEnable := True;
               IF #TSEND_C.DONE AND NOT #TSEND_C.BUSY THEN
                   #watchDogEnable := False;
                   #PingReqStep := 5;
               END_IF;
           5:
               IF #RcvDataNDR[13] AND #RcvDataNDLen[13] > 0 THEN
                   #PingReqStep := 6;
               END_IF;
           6:
               IF #RcvDataBuffer[13, 0] = 16#D0 AND #RcvDataBuffer[13, 1] = 16#00 THEN
                   #PingReqStep := 7;
               ELSE
                   #iError := True;
                   #iErrorID := 16#9040;
                   #ErrorSource := 16#13;
                   #PingReqStep := 8;
               END_IF;
           7:
               #PingRespCounter := #PingRespCounter + 1;
               #PingReqStep := 8;
           8:
               #RcvDataNDR[13] := False;
               #RcvDataNDLen[13] := 0;
               #PingReqStep := 0;
               #keepAliveEnable := False;
               #pinged := True;
       END_CASE;
   END_REGION ;
   REGION DISCONNET
       CASE #DisconnectStep OF
           0:
               ;
           1:
               #published := False;
               #subscribed := False;
               #unsubscribed := False;
               #pinged := False;
               #disconnected := False;
               #subscribedMsgReceived := False;
               #DisconnectStep := 2;
           2:
               #PingReqStep := 0;
               #TSENDATA[0] := 16#E0;
               #TSENDATA[1] := 16#00;
               #DisconnectStep := 3;
           3:
               #TSEND_C.LEN := 2;
               #watchDogEnable := False;
               #TSEND_C.REQ := True;
               #DisconnectStep := 4;
           4:
               IF #TSEND_C.DONE AND NOT #TSEND_C.BUSY THEN
                   #DisconnectStep := 5;
               END_IF;
           5:
               #MqttConnected := False;
               #watchDogEnable := False;
               #keepAliveEnable := False;
               #DisconnectStep := 0;
               #Enable := False;
               #disconnected := True;
       END_CASE;
   END_REGION ;
   REGION SubscribedMsgArrived
       IF (#RcvDataNDR[3] AND #RcvDataNDLen[3] > 0) AND NOT #p_trig[5] THEN
           #subscribedMsgIndex := 0;
           #RcvSubscribedMsgArrayIndex := 0;
           #SubscribedMsgRcvStep := 1;
       END_IF;
       #p_trig[5] := (#RcvDataNDR[3] AND #RcvDataNDLen[3] > 0);
       CASE #SubscribedMsgRcvStep OF
           0:
               ;
           1:
               #subscribedMsgReceived := False;
               #subscribedMsgQos.%X0 := #RcvDataBuffer[3, #subscribedMsgIndex].%X1;
               #subscribedMsgQos.%X1 := #RcvDataBuffer[3, #subscribedMsgIndex].%X2;
               IF #subscribedMsgQos >= 16#0 AND #subscribedMsgQos <= 16#2 THEN
                   #RLmultiplier := 1;
                   #subscribedPayloadDecodedRL := 0;
                   #RLencodedIndex := #subscribedMsgIndex + 1;
                   REPEAT
                       #RLencodedByte := #RcvDataBuffer[3, #RLencodedIndex];
                       #subscribedPayloadDecodedRL := #subscribedPayloadDecodedRL + (BYTE_TO_DINT(#RLencodedByte AND 127) * #RLmultiplier);
                       #RLmultiplier := #RLmultiplier * 128;
                       #RLencodedIndex := #RLencodedIndex + 1;
                       IF #RLmultiplier > 128 ** 3 THEN
                           #iError := False;
                           #iErrorID := 16#9050;
                           #ErrorSource := 16#0F;
                           #SubscribedMsgRcvStep := 30;
                       END_IF;
                   UNTIL (#RLencodedByte AND 128) = 0 END_REPEAT;
               ELSE
                   #iError := True;
                   #iErrorID := 16#9051;
                   #ErrorSource := 16#0F;
                   #SubscribedMsgRcvStep := 30;
               END_IF;
               #subscribedMsgIndex := #subscribedMsgIndex + 2;
               IF #subscribedPayloadDecodedRL >= 128 THEN
                   #subscribedMsgIndex := #subscribedMsgIndex + 1;
               END_IF;
               IF #subscribedPayloadDecodedRL >= 16384 THEN
                   #subscribedMsgIndex := #subscribedMsgIndex + 1;
               END_IF;
               IF #subscribedPayloadDecodedRL >= 2097152 THEN
                   #subscribedMsgIndex := #subscribedMsgIndex + 1;
               END_IF;
               #subscribedTopicLength_tmp.%B1 := #RcvDataBuffer[3, #subscribedMsgIndex];
               #subscribedTopicLength_tmp.%B0 := #RcvDataBuffer[3, #subscribedMsgIndex + 1];
               #subscribedTopicLength := WORD_TO_INT(#subscribedTopicLength_tmp);
               #subscribedMsgIndex := #subscribedMsgIndex + 2;
               #subscribedTopicNameIndex := #subscribedMsgIndex;
               #subscribedMsgIndex := #subscribedMsgIndex + #subscribedTopicLength;
               IF #subscribedMsgQos = 16#1 OR #subscribedMsgQos = 16#2 THEN
                   #subscribedPocketIdIndex := #subscribedMsgIndex;
                   #subscribedPayloadIndex := #subscribedMsgIndex + 2;
                   #subscribedMsgIndex := #subscribedMsgIndex + 2;
               ELSE
                   #subscribedPayloadIndex := #subscribedMsgIndex;
               END_IF;
               #subscribedPayloadLength := #subscribedPayloadDecodedRL - 2 - #subscribedTopicLength;
               IF #subscribedMsgQos = 16#1 OR #subscribedMsgQos = 16#2 THEN
                   #subscribedPayloadLength := #subscribedPayloadLength - 2;
                   #packetIdWordTmp.%B1 := #RcvDataBuffer[3, #subscribedPocketIdIndex];
                   #packetIdWordTmp.%B0 := #RcvDataBuffer[3, #subscribedPocketIdIndex + 1];
                   #TSENDATA[2] := #packetIdWordTmp.%B1;
                   #TSENDATA[3] := #packetIdWordTmp.%B0;
               END_IF;
               #SubscribedMsgRcvStep := 2;
           2:
               FOR #i := #RcvSubscribedMsgArrayIndex TO 9 DO
                   #ReceivedTopic[#i] := '';
                   #ReceivedMessage[#i] := '';
               END_FOR;
               IF #subscribedTopicLength > 254 THEN
                   #iError := True;
                   #iErrorID := 16#9054;
                   #ErrorSource := 16#0F;
                   #SubscribedMsgRcvStep := 30;
               END_IF;
               IF #subscribedPayloadLength > 254 THEN
                   #iError := True;
                   #iErrorID := 16#9055;
                   #ErrorSource := 16#0F;
                   #SubscribedMsgRcvStep := 30;
               END_IF;
               Chars_TO_Strg(Chars := #RcvDataBuffer[3],
                             pChars := #subscribedTopicNameIndex,
                             Cnt := INT_TO_UINT(#subscribedTopicLength),
                             Strg => #ReceivedTopic[#RcvSubscribedMsgArrayIndex]);
               Chars_TO_Strg(Chars := #RcvDataBuffer[3],
                             pChars := #subscribedPayloadIndex,
                             Cnt := DINT_TO_UINT(#subscribedPayloadLength),
                             Strg => #ReceivedMessage[#RcvSubscribedMsgArrayIndex]);
               #SubscribedMsgRcvStep := 3;
           3:
               #subscribedMsgReceived := True;
               #subscribedMsgIndex := #subscribedMsgIndex + DINT_TO_INT(#subscribedPayloadLength);
               CASE WORD_TO_INT(#subscribedMsgQos) OF
                   0:
                       #SubscribedMsgRcvStep := 24;
                   1:
                       #SubscribedMsgRcvStep := 20;
                   2:
                       #SubscribedMsgRcvStep := 10;
               END_CASE;
           10:
               #TSENDATA[0] := 16#50;
               #TSENDATA[1] := 16#02;
               #TSENDATA[2] := #packetIdWordTmp.%B1;
               #TSENDATA[3] := #packetIdWordTmp.%B0;
               #SubscribedMsgRcvStep := 11;
           11:
               UFILL_BLK(IN := 16#00,
                         COUNT := 255,
                         OUT => #RcvDataBuffer[7, 0]);
               #SubscribedMsgRcvStep := 12;
           12:
               #TSEND_C.LEN := 4;
               #RcvDataNDR[6] := False;
               #RcvDataNDLen[6] := 0;
               #TSEND_C.REQ := True;
               #SubscribedMsgRcvStep := 13;
           13:
               #watchDogEnable := True;
               IF #TSEND_C.DONE AND NOT #TSEND_C.BUSY THEN
                   #SubscribedMsgRcvStep := 14;
               END_IF;
           14:
               IF #RcvDataNDR[6] AND #RcvDataNDLen[6] > 0 THEN
                   #watchDogEnable := False;
                   IF #RcvDataBuffer[6, 0] = 16#62 AND #RcvDataBuffer[6, 1] = 16#02 THEN
                       #SubscribedMsgRcvStep := 15;
                   ELSE
                       #iError := True;
                       #iErrorID := 16#9052;
                       #ErrorSource := 16#06;
                       #SubscribedMsgRcvStep := 30;
                   END_IF;
               END_IF;
           15:
               IF #RcvDataBuffer[6, 2] = #packetIdWordTmp.%B1 AND #RcvDataBuffer[6, 3] = #packetIdWordTmp.%B0 THEN
                   #RcvDataNDR[6] := False;
                   #RcvDataNDLen[6] := 0;
                   #SubscribedMsgRcvStep := 16;
               ELSE
                   #iError := True;
                   #iErrorID := 16#9053;
                   #ErrorSource := 16#06;
                   #SubscribedMsgRcvStep := 30;
               END_IF;
           16:
               #TSENDATA[0] := 16#70;
               #TSENDATA[1] := 16#02;
               #TSENDATA[2] := #packetIdWordTmp.%B1;
               #TSENDATA[3] := #packetIdWordTmp.%B0;
               #SubscribedMsgRcvStep := 17;
           17:
               #TSEND_C.LEN := 4;
               #TSEND_C.REQ := True;
               #SubscribedMsgRcvStep := 18;
           18:
               #watchDogEnable := True;
               IF #TSEND_C.DONE AND NOT #TSEND_C.BUSY THEN
                   #watchDogEnable := False;
                   #SubscribedMsgRcvStep := 24;
               END_IF;
           20:
               #TSENDATA[0] := 16#40;
               #TSENDATA[1] := 16#02;
               #TSENDATA[2] := #packetIdWordTmp.%B1;
               #TSENDATA[3] := #packetIdWordTmp.%B0;
               #SubscribedMsgRcvStep := 21;
           21:
               #TSEND_C.LEN := 4;
               #TSEND_C.REQ := True;
               #SubscribedMsgRcvStep := 23;
           23:
               #watchDogEnable := True;
               IF #TSEND_C.DONE AND NOT #TSEND_C.BUSY THEN
                   #watchDogEnable := False;
                   #SubscribedMsgRcvStep := 24;
               END_IF;
           24:
               IF #subscribedMsgIndex < #RcvDataNDLen[3] THEN
                   #RcvSubscribedMsgArrayIndex := #RcvSubscribedMsgArrayIndex + 1;
                   #SubscribedMsgRcvStep := 1;
               ELSE
                   #SubscribedMsgRcvStep := 30;
               END_IF;
           30:
               UFILL_BLK(IN := 16#00,
                         COUNT := 255,
                         OUT => #RcvDataBuffer[3, 0]);
               FOR #i := 3 TO 7 DO
                   #RcvDataNDR[#i] := False;
                   #RcvDataNDLen[#i] := 0;
               END_FOR;
               #SubscribedMsgRcvStep := 0;
               #watchDogEnable := False;
       END_CASE;
   END_REGION ;
   REGION TIMERS
       #keepAliveTimerQ := #KeepAliveTimer.Q;
       #KeepAliveTimer(IN := #keepAliveEnable AND NOT #KeepAliveTimer.Q,
                       PT := #keepAliveTime);
       #WatchDogTimer(IN := #watchDogEnable AND (NOT #WatchDogTimer.Q),
                      PT := T#3s);
   END_REGION ;
   REGION Signal output
       #Busy := #Enable AND NOT #Idle;
       #Status.%X0 := #TcpConnected;
       #Status.%X1 := #MqttConnected;
       #Status.%X2 := #published;
       #Status.%X3 := #subscribed;
       #Status.%X4 := #unsubscribed;
       #Status.%X5 := #pinged;
       #Status.%X6 := #disconnected;
       #Status.%X7 := #subscribedMsgReceived;
       #Error := #iError;
       #ErrorID := #iErrorID;
   END_REGION ;
END_FUNCTION_BLOCK

// ===== library types =====

// folder: LMQTT

TYPE "LMQTT_typeConnParam"
TITLE = LMQTT_typeConnParams
// Specifies connection parameters for the mqtt connection
   STRUCT
      hwId : Hw_Any;   // Hardware identifier of the interface. 0: interface is selected automatically
      connId : Conn_Ouc;   // Unique connection identifier
      brokerAddress : Struct   // Information on the MQTT broker
         qdnAddress : String;   // Fully qualified domain name of the broker. must end with a dot "."
         ipAddress : IP_V4;   // If no FQDN is used, enter ip-address of the broker instead
         port : UInt;   // Enter the port of the mqtt broker
      END_STRUCT;
      tls : Struct   // Parameters for TLS encryption
         enableTls : Bool;   // TRUE: Enables TLS, FALSE: disable TLS
         validateServerIdentity : Bool;   // TRUE: Validate server certificate, FALSE: No validation of server certificate
         brokerCert : UDInt;   // ID of the broker's certificate in TIA Portal
         clientCert : UDInt;   // ID of the client's certificate in TIA Portal
      END_STRUCT;
      keepAlive : UInt;   // Keepalive mechanism for MQTT in seconds. 0: disabled.
   END_STRUCT;
END_TYPE

// folder: 01_Blocks/Utilities

